Universal Robots URScript: test_first_drawing_!.script

def Machining1():
  # Default parameters:
  global speed_ms = 0.3
  global speed_rads = 0.75
  global accel_mss = 3
  global accel_radss = 1.2
  global blend_radius_m = 0.001

  # Add subprograms here
  # Start of main program
  # Program generated by RoboDK v5.6.5 for UR10e on 02/02/2024 16:16:45
  # Using nominal kinematics.
  blend_radius_m = 0.001
  speed_ms = 1.000
  # set_reference(p[0.123734, -0.255000, -0.004586, 0.000000, 0.000000, 0.000000])
  set_tcp(p[0.000000, 0.000000, 0.252000, 0.000000, 0.000000, 0.000000])
  # Show Tool
  movej([-0.457372, -0.718365, -2.572418, -1.421607, 1.570796, 1.113424],accel_radss,speed_rads,0,blend_radius_m)
  movel([-0.457372, -0.718365, -2.572418, -1.421607, 1.570796, 1.113424],accel_mss,speed_ms,0,blend_radius_m)
  # Splitting Linear movement in 6 (instruction 7: MoveL 3)
  movel([-0.457372, -0.726970, -2.600418, -1.385001, 1.570796, 1.113424],accel_mss,speed_ms,0,blend_radius_m)
  movel([-0.457372, -0.737986, -2.628172, -1.346232, 1.570796, 1.113424],accel_mss,speed_ms,0,blend_radius_m)
  movel([-0.457372, -0.751770, -2.655662, -1.304957, 1.570796, 1.113424],accel_mss,speed_ms,0,blend_radius_m)
  movel([-0.457372, -0.768751, -2.682869, -1.260769, 1.570796, 1.113424],accel_mss,speed_ms,0,blend_radius_m)
  movel([-0.457372, -0.789449, -2.709765, -1.213175, 1.570796, 1.113424],accel_mss,speed_ms,0,blend_radius_m)
  movel([-0.457372, -0.814491, -2.736314, -1.161584, 1.570796, 1.113424],accel_mss,speed_ms,0,blend_radius_m)
  movel([-0.457372, -0.814491, -2.736314, -1.161584, 1.570796, 1.113424],accel_mss,speed_ms,0,blend_radius_m)
  speed_ms = 1.000
  movel([-0.457372, -0.814491, -2.736314, -1.161584, 1.570796, 1.113424],accel_mss,speed_ms,0,blend_radius_m)
  movel([-0.457372, -0.814491, -2.736314, -1.161584, 1.570796, 1.113424],accel_mss,speed_ms,0,blend_radius_m)
  movel([-0.457372, -0.814491, -2.736314, -1.161584, 1.570796, 1.113424],accel_mss,speed_ms,0,blend_radius_m)
  speed_ms = 0.005
  movel([-0.457372, -0.784984, -2.704412, -1.222993, 1.570796, 1.113424],accel_mss,speed_ms,0,blend_radius_m)
  speed_ms = 1.000
  movel([-0.457372, -0.814491, -2.736314, -1.161584, 1.570796, 1.113424],accel_mss,speed_ms,0,blend_radius_m)
  speed_ms = 0.040
  movel([-0.457372, -0.814491, -2.736314, -1.161584, 1.570796, 1.113424],accel_mss,speed_ms,0,blend_radius_m)
  speed_ms = 1.000
  movel([-0.457372, -0.814491, -2.736314, -1.161584, 1.570796, 1.113424],accel_mss,speed_ms,0,blend_radius_m)
  # Splitting Linear movement in 8 (instruction 21: MoveL 12)
  movel([-0.394298, -0.800154, -2.739094, -1.173141, 1.570796, 1.176498],accel_mss,speed_ms,0,blend_radius_m)
  movel([-0.332487, -0.789840, -2.741023, -1.181526, 1.570796, 1.238309],accel_mss,speed_ms,0,blend_radius_m)
  movel([-0.272464, -0.783804, -2.742125, -1.186460, 1.570796, 1.298332],accel_mss,speed_ms,0,blend_radius_m)
  movel([-0.214704, -0.782203, -2.742414, -1.187772, 1.570796, 1.356092],accel_mss,speed_ms,0,blend_radius_m)
  movel([-0.159605, -0.785077, -2.741894, -1.185418, 1.570796, 1.411192],accel_mss,speed_ms,0,blend_radius_m)
  movel([-0.107470, -0.792353, -2.740559, -1.179478, 1.570796, 1.463327],accel_mss,speed_ms,0,blend_radius_m)
  movel([-0.058503, -0.803844, -2.738390, -1.170155, 1.570796, 1.512293],accel_mss,speed_ms,0,blend_radius_m)
  movel([-0.012808, -0.819267, -2.735362, -1.157760, 1.570796, 1.557988],accel_mss,speed_ms,0,blend_radius_m)
  speed_ms = 0.005
  movel([-0.012808, -0.856350, -2.766620, -1.089418, 1.570796, 1.557988],accel_mss,speed_ms,0,blend_radius_m)
  speed_ms = 0.025
  movel([-0.015705, -0.866064, -2.764578, -1.081748, 1.570796, 1.555091],accel_mss,speed_ms,0,blend_radius_m)
  movel([-0.017368, -0.870976, -2.763523, -1.077890, 1.570796, 1.553429],accel_mss,speed_ms,0,blend_radius_m)
  movel([-0.019216, -0.875915, -2.762449, -1.074025, 1.570796, 1.551580],accel_mss,speed_ms,0,blend_radius_m)
  movel([-0.021279, -0.880866, -2.761357, -1.070166, 1.570796, 1.549518],accel_mss,speed_ms,0,blend_radius_m)
  movel([-0.023584, -0.885818, -2.760249, -1.066321, 1.570796, 1.547213],accel_mss,speed_ms,0,blend_radius_m)
  movel([-0.026163, -0.890765, -2.759128, -1.062496, 1.570796, 1.544633],accel_mss,speed_ms,0,blend_radius_m)
  movel([-0.029049, -0.895692, -2.757997, -1.058701, 1.570796, 1.541747],accel_mss,speed_ms,0,blend_radius_m)
  movel([-0.028017, -0.893565, -2.758487, -1.060337, 1.570796, 1.542779],accel_mss,speed_ms,0,blend_radius_m)
  movel([-0.027153, -0.890950, -2.759086, -1.062353, 1.570796, 1.543644],accel_mss,speed_ms,0,blend_radius_m)
  movel([-0.026737, -0.888547, -2.759633, -1.064209, 1.570796, 1.544059],accel_mss,speed_ms,0,blend_radius_m)
  movel([-0.026791, -0.887653, -2.759835, -1.064900, 1.570796, 1.544006],accel_mss,speed_ms,0,blend_radius_m)
  movel([-0.027063, -0.887078, -2.759965, -1.065346, 1.570796, 1.543734],accel_mss,speed_ms,0,blend_radius_m)
  movel([-0.027595, -0.886898, -2.760006, -1.065485, 1.570796, 1.543202],accel_mss,speed_ms,0,blend_radius_m)
  movel([-0.028284, -0.887183, -2.759942, -1.065264, 1.570796, 1.542513],accel_mss,speed_ms,0,blend_radius_m)
  movel([-0.029095, -0.887869, -2.759787, -1.064734, 1.570796, 1.541701],accel_mss,speed_ms,0,blend_radius_m)
  movel([-0.030017, -0.888906, -2.759551, -1.063932, 1.570796, 1.540780],accel_mss,speed_ms,0,blend_radius_m)
  movel([-0.032071, -0.891780, -2.758896, -1.061712, 1.570796, 1.538725],accel_mss,speed_ms,0,blend_radius_m)
  movel([-0.034255, -0.895333, -2.758079, -1.058976, 1.570796, 1.536542],accel_mss,speed_ms,0,blend_radius_m)
  movel([-0.038281, -0.902664, -2.756369, -1.053356, 1.570796, 1.532515],accel_mss,speed_ms,0,blend_radius_m)
  movel([-0.040683, -0.907306, -2.755268, -1.049815, 1.570796, 1.530113],accel_mss,speed_ms,0,blend_radius_m)
  movel([-0.044313, -0.913830, -2.753697, -1.044862, 1.570796, 1.526483],accel_mss,speed_ms,0,blend_radius_m)
  movel([-0.046379, -0.916993, -2.752926, -1.042470, 1.570796, 1.524417],accel_mss,speed_ms,0,blend_radius_m)
  movel([-0.048725, -0.920005, -2.752185, -1.040199, 1.570796, 1.522072],accel_mss,speed_ms,0,blend_radius_m)
  movel([-0.048271, -0.919131, -2.752401, -1.040857, 1.570796, 1.522525],accel_mss,speed_ms,0,blend_radius_m)
  movel([-0.048029, -0.917919, -2.752699, -1.041771, 1.570796, 1.522767],accel_mss,speed_ms,0,blend_radius_m)
  movel([-0.048062, -0.915005, -2.753411, -1.043973, 1.570796, 1.522735],accel_mss,speed_ms,0,blend_radius_m)
  movel([-0.048591, -0.912345, -2.754057, -1.045987, 1.570796, 1.522205],accel_mss,speed_ms,0,blend_radius_m)
  movel([-0.048976, -0.911448, -2.754274, -1.046667, 1.570796, 1.521820],accel_mss,speed_ms,0,blend_radius_m)
  movel([-0.049395, -0.911024, -2.754376, -1.046989, 1.570796, 1.521401],accel_mss,speed_ms,0,blend_radius_m)
  movel([-0.050483, -0.910927, -2.754399, -1.047062, 1.570796, 1.520313],accel_mss,speed_ms,0,blend_radius_m)
  movel([-0.051522, -0.911310, -2.754307, -1.046772, 1.570796, 1.519275],accel_mss,speed_ms,0,blend_radius_m)
  movel([-0.052515, -0.912075, -2.754122, -1.046192, 1.570796, 1.518281],accel_mss,speed_ms,0,blend_radius_m)
  movel([-0.053463, -0.913130, -2.753867, -1.045392, 1.570796, 1.517333],accel_mss,speed_ms,0,blend_radius_m)
  movel([-0.055213, -0.915686, -2.753245, -1.043458, 1.570796, 1.515583],accel_mss,speed_ms,0,blend_radius_m)
  movel([-0.056771, -0.918197, -2.752631, -1.041562, 1.570796, 1.514025],accel_mss,speed_ms,0,blend_radius_m)
  movel([-0.059370, -0.922009, -2.751689, -1.038691, 1.570796, 1.511427],accel_mss,speed_ms,0,blend_radius_m)
  movel([-0.062062, -0.925527, -2.750812, -1.036050, 1.570796, 1.508735],accel_mss,speed_ms,0,blend_radius_m)
  movel([-0.065029, -0.928771, -2.749996, -1.033622, 1.570796, 1.505768],accel_mss,speed_ms,0,blend_radius_m)
  movel([-0.068441, -0.931736, -2.749244, -1.031409, 1.570796, 1.502355],accel_mss,speed_ms,0,blend_radius_m)
  movel([-0.066682, -0.928859, -2.749974, -1.033557, 1.570796, 1.504114],accel_mss,speed_ms,0,blend_radius_m)
  movel([-0.065327, -0.925996, -2.750694, -1.035699, 1.570796, 1.505469],accel_mss,speed_ms,0,blend_radius_m)
  movel([-0.064965, -0.924615, -2.751040, -1.036734, 1.570796, 1.505831],accel_mss,speed_ms,0,blend_radius_m)
  movel([-0.064915, -0.923396, -2.751344, -1.037649, 1.570796, 1.505881],accel_mss,speed_ms,0,blend_radius_m)
  movel([-0.065209, -0.922449, -2.751580, -1.038360, 1.570796, 1.505588],accel_mss,speed_ms,0,blend_radius_m)
  movel([-0.065897, -0.921914, -2.751713, -1.038762, 1.570796, 1.504899],accel_mss,speed_ms,0,blend_radius_m)
  movel([-0.067234, -0.921954, -2.751703, -1.038732, 1.570796, 1.503563],accel_mss,speed_ms,0,blend_radius_m)
  movel([-0.068837, -0.922643, -2.751532, -1.038214, 1.570796, 1.501959],accel_mss,speed_ms,0,blend_radius_m)
  movel([-0.070570, -0.923760, -2.751254, -1.037376, 1.570796, 1.500226],accel_mss,speed_ms,0,blend_radius_m)
  movel([-0.072285, -0.925061, -2.750929, -1.036399, 1.570796, 1.498511],accel_mss,speed_ms,0,blend_radius_m)
  speed_ms = 0.005
  movel([-0.072285, -0.916497, -2.744962, -1.050930, 1.570796, 1.498511],accel_mss,speed_ms,0,blend_radius_m)
  speed_ms = 0.040
  movel([-0.064341, -0.944955, -2.737631, -1.029804, 1.570796, 1.506455],accel_mss,speed_ms,0,blend_radius_m)
  speed_ms = 0.005
  movel([-0.064341, -0.953673, -2.743494, -1.015222, 1.570796, 1.506455],accel_mss,speed_ms,0,blend_radius_m)
  speed_ms = 0.025
  movel([-0.063744, -0.951411, -2.744102, -1.016876, 1.570796, 1.507052],accel_mss,speed_ms,0,blend_radius_m)
  movel([-0.062886, -0.949058, -2.744731, -1.018600, 1.570796, 1.507911],accel_mss,speed_ms,0,blend_radius_m)
  movel([-0.061790, -0.946658, -2.745368, -1.020363, 1.570796, 1.509006],accel_mss,speed_ms,0,blend_radius_m)
  movel([-0.060471, -0.944238, -2.746007, -1.022144, 1.570796, 1.510325],accel_mss,speed_ms,0,blend_radius_m)
  movel([-0.058951, -0.941831, -2.746638, -1.023920, 1.570796, 1.511845],accel_mss,speed_ms,0,blend_radius_m)
  movel([-0.057246, -0.939476, -2.747252, -1.025660, 1.570796, 1.513550],accel_mss,speed_ms,0,blend_radius_m)
  movel([-0.055380, -0.937209, -2.747840, -1.027340, 1.570796, 1.515416],accel_mss,speed_ms,0,blend_radius_m)
  movel([-0.053368, -0.935059, -2.748394, -1.028936, 1.570796, 1.517428],accel_mss,speed_ms,0,blend_radius_m)
  movel([-0.050202, -0.932150, -2.749138, -1.031101, 1.570796, 1.520594],accel_mss,speed_ms,0,blend_radius_m)
  movel([-0.047049, -0.929750, -2.749748, -1.032891, 1.570796, 1.523747],accel_mss,speed_ms,0,blend_radius_m)
  movel([-0.043926, -0.927829, -2.750233, -1.034326, 1.570796, 1.526870],accel_mss,speed_ms,0,blend_radius_m)
  movel([-0.040855, -0.926363, -2.750602, -1.035424, 1.570796, 1.529941],accel_mss,speed_ms,0,blend_radius_m)
  movel([-0.037852, -0.925322, -2.750863, -1.036204, 1.570796, 1.532944],accel_mss,speed_ms,0,blend_radius_m)
  movel([-0.034930, -0.924675, -2.751025, -1.036689, 1.570796, 1.535866],accel_mss,speed_ms,0,blend_radius_m)
  movel([-0.032111, -0.924395, -2.751095, -1.036899, 1.570796, 1.538685],accel_mss,speed_ms,0,blend_radius_m)
  movel([-0.029407, -0.924448, -2.751082, -1.036859, 1.570796, 1.541389],accel_mss,speed_ms,0,blend_radius_m)
  movel([-0.026834, -0.924800, -2.750994, -1.036595, 1.570796, 1.543962],accel_mss,speed_ms,0,blend_radius_m)
  movel([-0.024404, -0.925419, -2.750839, -1.036131, 1.570796, 1.546392],accel_mss,speed_ms,0,blend_radius_m)
  movel([-0.020023, -0.927315, -2.750363, -1.034711, 1.570796, 1.550774],accel_mss,speed_ms,0,blend_radius_m)
  movel([-0.016359, -0.929848, -2.749723, -1.032818, 1.570796, 1.554437],accel_mss,speed_ms,0,blend_radius_m)
  movel([-0.013508, -0.932744, -2.748987, -1.030659, 1.570796, 1.557288],accel_mss,speed_ms,0,blend_radius_m)
  movel([-0.011055, -0.936237, -2.748091, -1.028061, 1.570796, 1.559741],accel_mss,speed_ms,0,blend_radius_m)
  movel([-0.009001, -0.940105, -2.747089, -1.025195, 1.570796, 1.561795],accel_mss,speed_ms,0,blend_radius_m)
  movel([-0.007301, -0.944288, -2.745994, -1.022107, 1.570796, 1.563495],accel_mss,speed_ms,0,blend_radius_m)
  movel([-0.005915, -0.948731, -2.744818, -1.018840, 1.570796, 1.564881],accel_mss,speed_ms,0,blend_radius_m)
  movel([-0.004799, -0.953378, -2.743573, -1.015438, 1.570796, 1.565997],accel_mss,speed_ms,0,blend_radius_m)
  movel([-0.003906, -0.958173, -2.742273, -1.011943, 1.570796, 1.566890],accel_mss,speed_ms,0,blend_radius_m)
  movel([-0.002624, -0.967997, -2.739559, -1.004833, 1.570796, 1.568172],accel_mss,speed_ms,0,blend_radius_m)
  movel([-0.001812, -0.974866, -2.737620, -0.999903, 1.570796, 1.568984],accel_mss,speed_ms,0,blend_radius_m)
  movel([-0.001114, -0.978051, -2.736709, -0.997629, 1.570796, 1.569682],accel_mss,speed_ms,0,blend_radius_m)
  movel([-0.000027, -0.980907, -2.735886, -0.995596, 1.570796, 1.570769],accel_mss,speed_ms,0,blend_radius_m)
  movel([0.001984, -0.984157, -2.734942, -0.993289, 1.570796, 1.572780],accel_mss,speed_ms,0,blend_radius_m)
  movel([0.003993, -0.987421, -2.733987, -0.990981, 1.570796, 1.574789],accel_mss,speed_ms,0,blend_radius_m)
  movel([0.004723, -0.989213, -2.733459, -0.989717, 1.570796, 1.575519],accel_mss,speed_ms,0,blend_radius_m)
  movel([0.005120, -0.991196, -2.732872, -0.988321, 1.570796, 1.575917],accel_mss,speed_ms,0,blend_radius_m)
  movel([0.005081, -0.993422, -2.732209, -0.986758, 1.570796, 1.575877],accel_mss,speed_ms,0,blend_radius_m)
  movel([0.004502, -0.995954, -2.731451, -0.984984, 1.570796, 1.575298],accel_mss,speed_ms,0,blend_radius_m)
  movel([0.006531, -0.989512, -2.733371, -0.989507, 1.570796, 1.577327],accel_mss,speed_ms,0,blend_radius_m)
  movel([0.008255, -0.983151, -2.735235, -0.994002, 1.570796, 1.579051],accel_mss,speed_ms,0,blend_radius_m)
  movel([0.011148, -0.970478, -2.738862, -1.003048, 1.570796, 1.581944],accel_mss,speed_ms,0,blend_radius_m)
  movel([0.012546, -0.963426, -2.740830, -1.008133, 1.570796, 1.583343],accel_mss,speed_ms,0,blend_radius_m)
  movel([0.013759, -0.956404, -2.742755, -1.013230, 1.570796, 1.584556],accel_mss,speed_ms,0,blend_radius_m)
  movel([0.015756, -0.942395, -2.746491, -1.023503, 1.570796, 1.586553],accel_mss,speed_ms,0,blend_radius_m)
  movel([0.017248, -0.928713, -2.750010, -1.033665, 1.570796, 1.588045],accel_mss,speed_ms,0,blend_radius_m)
  movel([0.017651, -0.921969, -2.751699, -1.038721, 1.570796, 1.588447],accel_mss,speed_ms,0,blend_radius_m)
  movel([0.017671, -0.915464, -2.753299, -1.043625, 1.570796, 1.588467],accel_mss,speed_ms,0,blend_radius_m)
  movel([0.017291, -0.910583, -2.754482, -1.047323, 1.570796, 1.588087],accel_mss,speed_ms,0,blend_radius_m)
  movel([0.016655, -0.905838, -2.755617, -1.050933, 1.570796, 1.587451],accel_mss,speed_ms,0,blend_radius_m)
  movel([0.016029, -0.901034, -2.756752, -1.054603, 1.570796, 1.586825],accel_mss,speed_ms,0,blend_radius_m)
  movel([0.015681, -0.895972, -2.757932, -1.058485, 1.570796, 1.586478],accel_mss,speed_ms,0,blend_radius_m)
  movel([0.015770, -0.894507, -2.758270, -1.059612, 1.570796, 1.586566],accel_mss,speed_ms,0,blend_radius_m)
  movel([0.016153, -0.892883, -2.758644, -1.060862, 1.570796, 1.586949],accel_mss,speed_ms,0,blend_radius_m)
  movel([0.016912, -0.891306, -2.759005, -1.062078, 1.570796, 1.587708],accel_mss,speed_ms,0,blend_radius_m)
  movel([0.017466, -0.890591, -2.759168, -1.062630, 1.570796, 1.588262],accel_mss,speed_ms,0,blend_radius_m)
  movel([0.018150, -0.889955, -2.759313, -1.063121, 1.570796, 1.588946],accel_mss,speed_ms,0,blend_radius_m)
  movel([0.019160, -0.889356, -2.759449, -1.063583, 1.570796, 1.589956],accel_mss,speed_ms,0,blend_radius_m)
  movel([0.020130, -0.889010, -2.759528, -1.063851, 1.570796, 1.590927],accel_mss,speed_ms,0,blend_radius_m)
  movel([0.025280, -0.887760, -2.759811, -1.064818, 1.570796, 1.596076],accel_mss,speed_ms,0,blend_radius_m)
  movel([0.029950, -0.887246, -2.759927, -1.065216, 1.570796, 1.600746],accel_mss,speed_ms,0,blend_radius_m)
  movel([0.034170, -0.887403, -2.759892, -1.065094, 1.570796, 1.604966],accel_mss,speed_ms,0,blend_radius_m)
  movel([0.037971, -0.888183, -2.759715, -1.064490, 1.570796, 1.608767],accel_mss,speed_ms,0,blend_radius_m)
  movel([0.041380, -0.889522, -2.759412, -1.063456, 1.570796, 1.612176],accel_mss,speed_ms,0,blend_radius_m)
  movel([0.044433, -0.891356, -2.758993, -1.062040, 1.570796, 1.615229],accel_mss,speed_ms,0,blend_radius_m)
  movel([0.047160, -0.893627, -2.758473, -1.060289, 1.570796, 1.617956],accel_mss,speed_ms,0,blend_radius_m)
  movel([0.049593, -0.896280, -2.757860, -1.058249, 1.570796, 1.620390],accel_mss,speed_ms,0,blend_radius_m)
  movel([0.051770, -0.899248, -2.757170, -1.055971, 1.570796, 1.622566],accel_mss,speed_ms,0,blend_radius_m)
  movel([0.053728, -0.902471, -2.756414, -1.053504, 1.570796, 1.624524],accel_mss,speed_ms,0,blend_radius_m)
  movel([0.057117, -0.909448, -2.754755, -1.048186, 1.570796, 1.627913],accel_mss,speed_ms,0,blend_radius_m)
  movel([0.062777, -0.923949, -2.751206, -1.037234, 1.570796, 1.633573],accel_mss,speed_ms,0,blend_radius_m)
  movel([0.063800, -0.926089, -2.750671, -1.035629, 1.570796, 1.634597],accel_mss,speed_ms,0,blend_radius_m)
  movel([0.064540, -0.926900, -2.750467, -1.035021, 1.570796, 1.635337],accel_mss,speed_ms,0,blend_radius_m)
  movel([0.065528, -0.927402, -2.750341, -1.034646, 1.570796, 1.636324],accel_mss,speed_ms,0,blend_radius_m)
  movel([0.067440, -0.927423, -2.750336, -1.034630, 1.570796, 1.638236],accel_mss,speed_ms,0,blend_radius_m)
  movel([0.068455, -0.927126, -2.750410, -1.034852, 1.570796, 1.639251],accel_mss,speed_ms,0,blend_radius_m)
  movel([0.069499, -0.926643, -2.750532, -1.035214, 1.570796, 1.640295],accel_mss,speed_ms,0,blend_radius_m)
  movel([0.071627, -0.925216, -2.750890, -1.036283, 1.570796, 1.642424],accel_mss,speed_ms,0,blend_radius_m)
  movel([0.073755, -0.923294, -2.751370, -1.037725, 1.570796, 1.644551],accel_mss,speed_ms,0,blend_radius_m)
  movel([0.075801, -0.921041, -2.751929, -1.039419, 1.570796, 1.646597],accel_mss,speed_ms,0,blend_radius_m)
  movel([0.077686, -0.918613, -2.752528, -1.041247, 1.570796, 1.648483],accel_mss,speed_ms,0,blend_radius_m)
  movel([0.079336, -0.916165, -2.753128, -1.043095, 1.570796, 1.650133],accel_mss,speed_ms,0,blend_radius_m)
  movel([0.080656, -0.913866, -2.753688, -1.044834, 1.570796, 1.651452],accel_mss,speed_ms,0,blend_radius_m)
  movel([0.082630, -0.909930, -2.754640, -1.047820, 1.570796, 1.653426],accel_mss,speed_ms,0,blend_radius_m)
  movel([0.084460, -0.905965, -2.755587, -1.050837, 1.570796, 1.655256],accel_mss,speed_ms,0,blend_radius_m)
  movel([0.087673, -0.898016, -2.757457, -1.056916, 1.570796, 1.658469],accel_mss,speed_ms,0,blend_radius_m)
  movel([0.090296, -0.890146, -2.759269, -1.062974, 1.570796, 1.661093],accel_mss,speed_ms,0,blend_radius_m)
  movel([0.092317, -0.882486, -2.760996, -1.068906, 1.570796, 1.663113],accel_mss,speed_ms,0,blend_radius_m)
  movel([0.092972, -0.879636, -2.761629, -1.071123, 1.570796, 1.663768],accel_mss,speed_ms,0,blend_radius_m)
  movel([0.093861, -0.876714, -2.762274, -1.073401, 1.570796, 1.664657],accel_mss,speed_ms,0,blend_radius_m)
  movel([0.094496, -0.875233, -2.762598, -1.074558, 1.570796, 1.665293],accel_mss,speed_ms,0,blend_radius_m)
  movel([0.095316, -0.873730, -2.762926, -1.075733, 1.570796, 1.666112],accel_mss,speed_ms,0,blend_radius_m)
  movel([0.096359, -0.872215, -2.763255, -1.076919, 1.570796, 1.667155],accel_mss,speed_ms,0,blend_radius_m)
  movel([0.097667, -0.870690, -2.763585, -1.078114, 1.570796, 1.668463],accel_mss,speed_ms,0,blend_radius_m)
  movel([0.099645, -0.869011, -2.763947, -1.079431, 1.570796, 1.670442],accel_mss,speed_ms,0,blend_radius_m)
  movel([0.101657, -0.867976, -2.764169, -1.080244, 1.570796, 1.672454],accel_mss,speed_ms,0,blend_radius_m)
  movel([0.103554, -0.867531, -2.764264, -1.080594, 1.570796, 1.674351],accel_mss,speed_ms,0,blend_radius_m)
  movel([0.105201, -0.867609, -2.764248, -1.080532, 1.570796, 1.675998],accel_mss,speed_ms,0,blend_radius_m)
  movel([0.107545, -0.868375, -2.764083, -1.079931, 1.570796, 1.678341],accel_mss,speed_ms,0,blend_radius_m)
  movel([0.109640, -0.869541, -2.763833, -1.079015, 1.570796, 1.680436],accel_mss,speed_ms,0,blend_radius_m)
  movel([0.113241, -0.872557, -2.763181, -1.076651, 1.570796, 1.684037],accel_mss,speed_ms,0,blend_radius_m)
  movel([0.114694, -0.874237, -2.762816, -1.075336, 1.570796, 1.685491],accel_mss,speed_ms,0,blend_radius_m)
  movel([0.115871, -0.876122, -2.762404, -1.073864, 1.570796, 1.686668],accel_mss,speed_ms,0,blend_radius_m)
  movel([0.116792, -0.878190, -2.761949, -1.072250, 1.570796, 1.687588],accel_mss,speed_ms,0,blend_radius_m)
  movel([0.117465, -0.880433, -2.761453, -1.070503, 1.570796, 1.688262],accel_mss,speed_ms,0,blend_radius_m)
  movel([0.117909, -0.882834, -2.760919, -1.068636, 1.570796, 1.688705],accel_mss,speed_ms,0,blend_radius_m)
  movel([0.118158, -0.888067, -2.759742, -1.064581, 1.570796, 1.688954],accel_mss,speed_ms,0,blend_radius_m)
  movel([0.117990, -0.890869, -2.759105, -1.062415, 1.570796, 1.688786],accel_mss,speed_ms,0,blend_radius_m)
  movel([0.117154, -0.896775, -2.757746, -1.057869, 1.570796, 1.687950],accel_mss,speed_ms,0,blend_radius_m)
  movel([0.115733, -0.903003, -2.756289, -1.053097, 1.570796, 1.686529],accel_mss,speed_ms,0,blend_radius_m)
  movel([0.113833, -0.909462, -2.754752, -1.048175, 1.570796, 1.684629],accel_mss,speed_ms,0,blend_radius_m)
  movel([0.111569, -0.916046, -2.753158, -1.043186, 1.570796, 1.682366],accel_mss,speed_ms,0,blend_radius_m)
  movel([0.107783, -0.925727, -2.750762, -1.035900, 1.570796, 1.678579],accel_mss,speed_ms,0,blend_radius_m)
  movel([0.105653, -0.930585, -2.749536, -1.032268, 1.570796, 1.676449],accel_mss,speed_ms,0,blend_radius_m)
  movel([0.103334, -0.935430, -2.748298, -1.028661, 1.570796, 1.674131],accel_mss,speed_ms,0,blend_radius_m)
  movel([0.100810, -0.940237, -2.747054, -1.025097, 1.570796, 1.671606],accel_mss,speed_ms,0,blend_radius_m)
  movel([0.098064, -0.944987, -2.745810, -1.021592, 1.570796, 1.668860],accel_mss,speed_ms,0,blend_radius_m)
  movel([0.095066, -0.949669, -2.744568, -1.018152, 1.570796, 1.665862],accel_mss,speed_ms,0,blend_radius_m)
  movel([0.091805, -0.954256, -2.743336, -1.014797, 1.570796, 1.662601],accel_mss,speed_ms,0,blend_radius_m)
  movel([0.086890, -0.960481, -2.741642, -1.010267, 1.570796, 1.657687],accel_mss,speed_ms,0,blend_radius_m)
  movel([0.084158, -0.963622, -2.740776, -1.007991, 1.570796, 1.654954],accel_mss,speed_ms,0,blend_radius_m)
  movel([0.081297, -0.966623, -2.739942, -1.005824, 1.570796, 1.652094],accel_mss,speed_ms,0,blend_radius_m)
  movel([0.078356, -0.969360, -2.739177, -1.003852, 1.570796, 1.649152],accel_mss,speed_ms,0,blend_radius_m)
  movel([0.075374, -0.971717, -2.738513, -1.002159, 1.570796, 1.646170],accel_mss,speed_ms,0,blend_radius_m)
  movel([0.072391, -0.973574, -2.737987, -1.000828, 1.570796, 1.643187],accel_mss,speed_ms,0,blend_radius_m)
  movel([0.070913, -0.974281, -2.737786, -1.000322, 1.570796, 1.641710],accel_mss,speed_ms,0,blend_radius_m)
  movel([0.069453, -0.974815, -2.737634, -0.999940, 1.570796, 1.640249],accel_mss,speed_ms,0,blend_radius_m)
  movel([0.067859, -0.975193, -2.737527, -0.999670, 1.570796, 1.638655],accel_mss,speed_ms,0,blend_radius_m)
  movel([0.066391, -0.975318, -2.737491, -0.999580, 1.570796, 1.637187],accel_mss,speed_ms,0,blend_radius_m)
  movel([0.065038, -0.975217, -2.737520, -0.999652, 1.570796, 1.635834],accel_mss,speed_ms,0,blend_radius_m)
  movel([0.063796, -0.974907, -2.737608, -0.999874, 1.570796, 1.634592],accel_mss,speed_ms,0,blend_radius_m)
  movel([0.061607, -0.973759, -2.737935, -1.000696, 1.570796, 1.632403],accel_mss,speed_ms,0,blend_radius_m)
  movel([0.059773, -0.972041, -2.738421, -1.001927, 1.570796, 1.630570],accel_mss,speed_ms,0,blend_radius_m)
  movel([0.058238, -0.969934, -2.739015, -1.003440, 1.570796, 1.629034],accel_mss,speed_ms,0,blend_radius_m)
  movel([0.056949, -0.967612, -2.739666, -1.005111, 1.570796, 1.627745],accel_mss,speed_ms,0,blend_radius_m)
  movel([0.054905, -0.963026, -2.740941, -1.008422, 1.570796, 1.625701],accel_mss,speed_ms,0,blend_radius_m)
  movel([0.053979, -0.960865, -2.741536, -1.009988, 1.570796, 1.624775],accel_mss,speed_ms,0,blend_radius_m)
  movel([0.052794, -0.958972, -2.742055, -1.011362, 1.570796, 1.623591],accel_mss,speed_ms,0,blend_radius_m)
  movel([0.051998, -0.958284, -2.742243, -1.011862, 1.570796, 1.622794],accel_mss,speed_ms,0,blend_radius_m)
  movel([0.051005, -0.957852, -2.742361, -1.012176, 1.570796, 1.621801],accel_mss,speed_ms,0,blend_radius_m)
  movel([0.049778, -0.957741, -2.742391, -1.012257, 1.570796, 1.620574],accel_mss,speed_ms,0,blend_radius_m)
  movel([0.048272, -0.958009, -2.742318, -1.012062, 1.570796, 1.619069],accel_mss,speed_ms,0,blend_radius_m)
  movel([0.048603, -0.958015, -2.742316, -1.012058, 1.570796, 1.619399],accel_mss,speed_ms,0,blend_radius_m)
  movel([0.048805, -0.958251, -2.742252, -1.011886, 1.570796, 1.619602],accel_mss,speed_ms,0,blend_radius_m)
  movel([0.048847, -0.959360, -2.741949, -1.011080, 1.570796, 1.619643],accel_mss,speed_ms,0,blend_radius_m)
  movel([0.048450, -0.961220, -2.741439, -1.009731, 1.570796, 1.619246],accel_mss,speed_ms,0,blend_radius_m)
  movel([0.047686, -0.963709, -2.740752, -1.007928, 1.570796, 1.618482],accel_mss,speed_ms,0,blend_radius_m)
  movel([0.045299, -0.970090, -2.738971, -1.003327, 1.570796, 1.616095],accel_mss,speed_ms,0,blend_radius_m)
  movel([0.042178, -0.977549, -2.736853, -0.997987, 1.570796, 1.612974],accel_mss,speed_ms,0,blend_radius_m)
  movel([0.035644, -0.992051, -2.732618, -0.987721, 1.570796, 1.606440],accel_mss,speed_ms,0,blend_radius_m)
  movel([0.031683, -1.000255, -2.730152, -0.981982, 1.570796, 1.602480],accel_mss,speed_ms,0,blend_radius_m)
  movel([0.026965, -1.008739, -2.727549, -0.976102, 1.570796, 1.597761],accel_mss,speed_ms,0,blend_radius_m)
  movel([0.022176, -1.017023, -2.724953, -0.970413, 1.570796, 1.592972],accel_mss,speed_ms,0,blend_radius_m)
  movel([0.017300, -1.025189, -2.722341, -0.964859, 1.570796, 1.588096],accel_mss,speed_ms,0,blend_radius_m)
  movel([0.007614, -1.040765, -2.717211, -0.954413, 1.570796, 1.578410],accel_mss,speed_ms,0,blend_radius_m)
  movel([0.002683, -1.048049, -2.714744, -0.949595, 1.570796, 1.573479],accel_mss,speed_ms,0,blend_radius_m)
  movel([0.000072, -1.051561, -2.713539, -0.947289, 1.570796, 1.570868],accel_mss,speed_ms,0,blend_radius_m)
  movel([-0.002659, -1.054953, -2.712365, -0.945071, 1.570796, 1.568137],accel_mss,speed_ms,0,blend_radius_m)
  movel([-0.005542, -1.058200, -2.711233, -0.942956, 1.570796, 1.565254],accel_mss,speed_ms,0,blend_radius_m)
  movel([-0.008588, -1.061277, -2.710151, -0.940961, 1.570796, 1.562208],accel_mss,speed_ms,0,blend_radius_m)
  movel([-0.008300, -1.055649, -2.712123, -0.944617, 1.570796, 1.562497],accel_mss,speed_ms,0,blend_radius_m)
  movel([-0.008450, -1.054105, -2.712660, -0.945624, 1.570796, 1.562346],accel_mss,speed_ms,0,blend_radius_m)
  movel([-0.008799, -1.053604, -2.712833, -0.945952, 1.570796, 1.561997],accel_mss,speed_ms,0,blend_radius_m)
  movel([-0.009432, -1.053476, -2.712878, -0.946035, 1.570796, 1.561364],accel_mss,speed_ms,0,blend_radius_m)
  movel([-0.010104, -1.053708, -2.712797, -0.945883, 1.570796, 1.560692],accel_mss,speed_ms,0,blend_radius_m)
  movel([-0.010802, -1.054169, -2.712638, -0.945583, 1.570796, 1.559994],accel_mss,speed_ms,0,blend_radius_m)
  movel([-0.014070, -1.056982, -2.711659, -0.943748, 1.570796, 1.556726],accel_mss,speed_ms,0,blend_radius_m)
  movel([-0.016026, -1.058338, -2.711184, -0.942867, 1.570796, 1.554770],accel_mss,speed_ms,0,blend_radius_m)
  movel([-0.018005, -1.059430, -2.710801, -0.942158, 1.570796, 1.552792],accel_mss,speed_ms,0,blend_radius_m)
  movel([-0.019956, -1.060230, -2.710520, -0.941639, 1.570796, 1.550841],accel_mss,speed_ms,0,blend_radius_m)
  movel([-0.020553, -1.060316, -2.710490, -0.941583, 1.570796, 1.550244],accel_mss,speed_ms,0,blend_radius_m)
  movel([-0.020750, -1.060021, -2.710594, -0.941775, 1.570796, 1.550047],accel_mss,speed_ms,0,blend_radius_m)
  movel([-0.020330, -1.058298, -2.711198, -0.942893, 1.570796, 1.550466],accel_mss,speed_ms,0,blend_radius_m)
  movel([-0.020427, -1.057821, -2.711365, -0.943202, 1.570796, 1.550369],accel_mss,speed_ms,0,blend_radius_m)
  movel([-0.020779, -1.057569, -2.711454, -0.943367, 1.570796, 1.550018],accel_mss,speed_ms,0,blend_radius_m)
  movel([-0.021298, -1.057529, -2.711467, -0.943393, 1.570796, 1.549498],accel_mss,speed_ms,0,blend_radius_m)
  movel([-0.021902, -1.057693, -2.711410, -0.943286, 1.570796, 1.548894],accel_mss,speed_ms,0,blend_radius_m)
  movel([-0.023143, -1.058460, -2.711142, -0.942788, 1.570796, 1.547654],accel_mss,speed_ms,0,blend_radius_m)
  movel([-0.031654, -1.066064, -2.708452, -0.937873, 1.570796, 1.539142],accel_mss,speed_ms,0,blend_radius_m)
  movel([-0.029187, -1.063378, -2.709408, -0.939603, 1.570796, 1.541609],accel_mss,speed_ms,0,blend_radius_m)
  movel([-0.026775, -1.060512, -2.710421, -0.941457, 1.570796, 1.544022],accel_mss,speed_ms,0,blend_radius_m)
  movel([-0.024437, -1.057512, -2.711473, -0.943404, 1.570796, 1.546359],accel_mss,speed_ms,0,blend_radius_m)
  movel([-0.022179, -1.054410, -2.712554, -0.945425, 1.570796, 1.548617],accel_mss,speed_ms,0,blend_radius_m)
  movel([-0.017959, -1.048048, -2.714745, -0.949597, 1.570796, 1.552837],accel_mss,speed_ms,0,blend_radius_m)
  movel([-0.014223, -1.041744, -2.716882, -0.953763, 1.570796, 1.556573],accel_mss,speed_ms,0,blend_radius_m)
  movel([-0.010453, -1.034858, -2.719180, -0.958352, 1.570796, 1.560343],accel_mss,speed_ms,0,blend_radius_m)
  movel([-0.006899, -1.027854, -2.721477, -0.963057, 1.570796, 1.563897],accel_mss,speed_ms,0,blend_radius_m)
  movel([-0.005272, -1.024335, -2.722617, -0.965438, 1.570796, 1.565524],accel_mss,speed_ms,0,blend_radius_m)
  movel([-0.003775, -1.020815, -2.723747, -0.967828, 1.570796, 1.567021],accel_mss,speed_ms,0,blend_radius_m)
  movel([-0.002443, -1.017311, -2.724861, -0.970216, 1.570796, 1.568354],accel_mss,speed_ms,0,blend_radius_m)
  movel([-0.001298, -1.013828, -2.725960, -0.972601, 1.570796, 1.569498],accel_mss,speed_ms,0,blend_radius_m)
  movel([-0.000737, -1.011694, -2.726629, -0.974066, 1.570796, 1.570060],accel_mss,speed_ms,0,blend_radius_m)
  movel([-0.000345, -1.009600, -2.727281, -0.975507, 1.570796, 1.570452],accel_mss,speed_ms,0,blend_radius_m)
  movel([-0.000026, -1.005553, -2.728533, -0.978303, 1.570796, 1.570770],accel_mss,speed_ms,0,blend_radius_m)
  movel([-0.000280, -1.001733, -2.729702, -0.980953, 1.570796, 1.570517],accel_mss,speed_ms,0,blend_radius_m)
  movel([-0.001044, -0.998182, -2.730780, -0.983427, 1.570796, 1.569752],accel_mss,speed_ms,0,blend_radius_m)
  movel([-0.002245, -0.994936, -2.731756, -0.985696, 1.570796, 1.568551],accel_mss,speed_ms,0,blend_radius_m)
  movel([-0.003811, -0.992035, -2.732623, -0.987732, 1.570796, 1.566986],accel_mss,speed_ms,0,blend_radius_m)
  movel([-0.005678, -0.989521, -2.733368, -0.989500, 1.570796, 1.565118],accel_mss,speed_ms,0,blend_radius_m)
  movel([-0.007767, -0.987427, -2.733985, -0.990977, 1.570796, 1.563029],accel_mss,speed_ms,0,blend_radius_m)
  movel([-0.009278, -0.986640, -2.734216, -0.991533, 1.570796, 1.561518],accel_mss,speed_ms,0,blend_radius_m)
  movel([-0.011068, -0.986527, -2.734249, -0.991612, 1.570796, 1.559729],accel_mss,speed_ms,0,blend_radius_m)
  movel([-0.013033, -0.987029, -2.734102, -0.991258, 1.570796, 1.557763],accel_mss,speed_ms,0,blend_radius_m)
  movel([-0.015068, -0.988082, -2.733793, -0.990515, 1.570796, 1.555729],accel_mss,speed_ms,0,blend_radius_m)
  movel([-0.017075, -0.989619, -2.733339, -0.989431, 1.570796, 1.553721],accel_mss,speed_ms,0,blend_radius_m)
  movel([-0.018953, -0.991579, -2.732758, -0.988052, 1.570796, 1.551843],accel_mss,speed_ms,0,blend_radius_m)
  movel([-0.020593, -0.993887, -2.732070, -0.986432, 1.570796, 1.550204],accel_mss,speed_ms,0,blend_radius_m)
  movel([-0.021902, -0.996480, -2.731293, -0.984616, 1.570796, 1.548895],accel_mss,speed_ms,0,blend_radius_m)
  movel([-0.023588, -1.000418, -2.730103, -0.981868, 1.570796, 1.547208],accel_mss,speed_ms,0,blend_radius_m)
  movel([-0.025438, -1.004334, -2.728907, -0.979148, 1.570796, 1.545359],accel_mss,speed_ms,0,blend_radius_m)
  movel([-0.027473, -1.008197, -2.727717, -0.976475, 1.570796, 1.543323],accel_mss,speed_ms,0,blend_radius_m)
  movel([-0.029724, -1.011987, -2.726537, -0.973865, 1.570796, 1.541072],accel_mss,speed_ms,0,blend_radius_m)
  movel([-0.032206, -1.015673, -2.725380, -0.971337, 1.570796, 1.538590],accel_mss,speed_ms,0,blend_radius_m)
  movel([-0.034949, -1.019235, -2.724251, -0.968904, 1.570796, 1.535847],accel_mss,speed_ms,0,blend_radius_m)
  movel([-0.037977, -1.022651, -2.723158, -0.966579, 1.570796, 1.532820],accel_mss,speed_ms,0,blend_radius_m)
  movel([-0.041308, -1.025896, -2.722112, -0.964381, 1.570796, 1.529489],accel_mss,speed_ms,0,blend_radius_m)
  movel([-0.043141, -1.027404, -2.721623, -0.963361, 1.570796, 1.527656],accel_mss,speed_ms,0,blend_radius_m)
  movel([-0.045025, -1.028711, -2.721198, -0.962480, 1.570796, 1.525771],accel_mss,speed_ms,0,blend_radius_m)
  movel([-0.048851, -1.030951, -2.720466, -0.960972, 1.570796, 1.521945],accel_mss,speed_ms,0,blend_radius_m)
  movel([-0.051855, -1.032427, -2.719982, -0.959980, 1.570796, 1.518942],accel_mss,speed_ms,0,blend_radius_m)
  movel([-0.054729, -1.033492, -2.719631, -0.959266, 1.570796, 1.516067],accel_mss,speed_ms,0,blend_radius_m)
  movel([-0.057472, -1.034176, -2.719405, -0.958808, 1.570796, 1.513324],accel_mss,speed_ms,0,blend_radius_m)
  movel([-0.060093, -1.034512, -2.719294, -0.958583, 1.570796, 1.510703],accel_mss,speed_ms,0,blend_radius_m)
  movel([-0.062595, -1.034534, -2.719287, -0.958568, 1.570796, 1.508201],accel_mss,speed_ms,0,blend_radius_m)
  movel([-0.064982, -1.034272, -2.719374, -0.958744, 1.570796, 1.505814],accel_mss,speed_ms,0,blend_radius_m)
  movel([-0.067250, -1.033750, -2.719546, -0.959093, 1.570796, 1.503546],accel_mss,speed_ms,0,blend_radius_m)
  movel([-0.069405, -1.033003, -2.719792, -0.959594, 1.570796, 1.501391],accel_mss,speed_ms,0,blend_radius_m)
  movel([-0.071449, -1.032061, -2.720102, -0.960226, 1.570796, 1.499347],accel_mss,speed_ms,0,blend_radius_m)
  movel([-0.073381, -1.030945, -2.720468, -0.960975, 1.570796, 1.497415],accel_mss,speed_ms,0,blend_radius_m)
  movel([-0.076913, -1.028330, -2.721322, -0.962736, 1.570796, 1.493884],accel_mss,speed_ms,0,blend_radius_m)
  movel([-0.080004, -1.025382, -2.722279, -0.964728, 1.570796, 1.490792],accel_mss,speed_ms,0,blend_radius_m)
  movel([-0.082651, -1.022337, -2.723259, -0.966793, 1.570796, 1.488146],accel_mss,speed_ms,0,blend_radius_m)
  movel([-0.084495, -1.019837, -2.724059, -0.968493, 1.570796, 1.486301],accel_mss,speed_ms,0,blend_radius_m)
  movel([-0.086208, -1.017088, -2.724932, -0.970369, 1.570796, 1.484589],accel_mss,speed_ms,0,blend_radius_m)
  movel([-0.087768, -1.014096, -2.725876, -0.972417, 1.570796, 1.483028],accel_mss,speed_ms,0,blend_radius_m)
  movel([-0.089137, -1.010871, -2.726886, -0.974632, 1.570796, 1.481659],accel_mss,speed_ms,0,blend_radius_m)
  movel([-0.090297, -1.007423, -2.727956, -0.977010, 1.570796, 1.480500],accel_mss,speed_ms,0,blend_radius_m)
  movel([-0.091211, -1.003760, -2.729083, -0.979546, 1.570796, 1.479586],accel_mss,speed_ms,0,blend_radius_m)
  movel([-0.091847, -0.999887, -2.730264, -0.982238, 1.570796, 1.478949],accel_mss,speed_ms,0,blend_radius_m)
  movel([-0.092176, -0.995812, -2.731494, -0.985083, 1.570796, 1.478621],accel_mss,speed_ms,0,blend_radius_m)
  movel([-0.092167, -0.991541, -2.732769, -0.988079, 1.570796, 1.478629],accel_mss,speed_ms,0,blend_radius_m)
  movel([-0.091786, -0.987087, -2.734085, -0.991217, 1.570796, 1.479010],accel_mss,speed_ms,0,blend_radius_m)
  movel([-0.091001, -0.982448, -2.735440, -0.994501, 1.570796, 1.479795],accel_mss,speed_ms,0,blend_radius_m)
  movel([-0.089771, -0.977635, -2.736828, -0.997926, 1.570796, 1.481025],accel_mss,speed_ms,0,blend_radius_m)
  movel([-0.088067, -0.972657, -2.738247, -1.001485, 1.570796, 1.482729],accel_mss,speed_ms,0,blend_radius_m)
  movel([-0.085849, -0.967515, -2.739693, -1.005180, 1.570796, 1.484947],accel_mss,speed_ms,0,blend_radius_m)
  movel([-0.083084, -0.962228, -2.741161, -1.009000, 1.570796, 1.487712],accel_mss,speed_ms,0,blend_radius_m)
  movel([-0.079736, -0.956800, -2.742647, -1.012942, 1.570796, 1.491060],accel_mss,speed_ms,0,blend_radius_m)
  movel([-0.078244, -0.954732, -2.743208, -1.014449, 1.570796, 1.492552],accel_mss,speed_ms,0,blend_radius_m)
  movel([-0.077402, -0.953783, -2.743464, -1.015142, 1.570796, 1.493394],accel_mss,speed_ms,0,blend_radius_m)
  movel([-0.076483, -0.952964, -2.743685, -1.015741, 1.570796, 1.494314],accel_mss,speed_ms,0,blend_radius_m)
  movel([-0.075051, -0.952139, -2.743907, -1.016344, 1.570796, 1.495745],accel_mss,speed_ms,0,blend_radius_m)
  movel([-0.073726, -0.951837, -2.743988, -1.016564, 1.570796, 1.497071],accel_mss,speed_ms,0,blend_radius_m)
  movel([-0.072569, -0.951977, -2.743950, -1.016462, 1.570796, 1.498227],accel_mss,speed_ms,0,blend_radius_m)
  movel([-0.071650, -0.952476, -2.743816, -1.016097, 1.570796, 1.499146],accel_mss,speed_ms,0,blend_radius_m)
  movel([-0.070227, -0.954257, -2.743336, -1.014796, 1.570796, 1.500570],accel_mss,speed_ms,0,blend_radius_m)
  movel([-0.069296, -0.956555, -2.742713, -1.013120, 1.570796, 1.501500],accel_mss,speed_ms,0,blend_radius_m)
  movel([-0.067994, -0.961593, -2.741336, -1.009460, 1.570796, 1.502802],accel_mss,speed_ms,0,blend_radius_m)
  movel([-0.067482, -0.962340, -2.741130, -1.008919, 1.570796, 1.503314],accel_mss,speed_ms,0,blend_radius_m)
  movel([-0.067015, -0.962322, -2.741135, -1.008932, 1.570796, 1.503782],accel_mss,speed_ms,0,blend_radius_m)
  movel([-0.066333, -0.961956, -2.741236, -1.009197, 1.570796, 1.504463],accel_mss,speed_ms,0,blend_radius_m)
  movel([-0.065449, -0.959415, -2.741934, -1.011041, 1.570796, 1.505347],accel_mss,speed_ms,0,blend_radius_m)
  movel([-0.064723, -0.956867, -2.742629, -1.012893, 1.570796, 1.506074],accel_mss,speed_ms,0,blend_radius_m)
  movel([-0.063159, -0.964473, -2.740540, -1.007376, 1.570796, 1.507637],accel_mss,speed_ms,0,blend_radius_m)
  movel([-0.061322, -0.971801, -2.738489, -1.002099, 1.570796, 1.509475],accel_mss,speed_ms,0,blend_radius_m)
  movel([-0.059217, -0.978853, -2.736479, -0.997057, 1.570796, 1.511580],accel_mss,speed_ms,0,blend_radius_m)
  movel([-0.056851, -0.985636, -2.734510, -0.992243, 1.570796, 1.513946],accel_mss,speed_ms,0,blend_radius_m)
  movel([-0.055705, -0.988480, -2.733675, -0.990234, 1.570796, 1.515091],accel_mss,speed_ms,0,blend_radius_m)
  movel([-0.054214, -0.991193, -2.732873, -0.988323, 1.570796, 1.516582],accel_mss,speed_ms,0,blend_radius_m)
  movel([-0.053288, -0.992366, -2.732524, -0.987499, 1.570796, 1.517508],accel_mss,speed_ms,0,blend_radius_m)
  movel([-0.052214, -0.993345, -2.732232, -0.986812, 1.570796, 1.518582],accel_mss,speed_ms,0,blend_radius_m)
  movel([-0.050968, -0.994073, -2.732015, -0.986301, 1.570796, 1.519828],accel_mss,speed_ms,0,blend_radius_m)
  movel([-0.049530, -0.994493, -2.731889, -0.986007, 1.570796, 1.521266],accel_mss,speed_ms,0,blend_radius_m)
  movel([-0.048410, -0.994565, -2.731868, -0.985957, 1.570796, 1.522386],accel_mss,speed_ms,0,blend_radius_m)
  movel([-0.045989, -0.994112, -2.732003, -0.986274, 1.570796, 1.524807],accel_mss,speed_ms,0,blend_radius_m)
  movel([-0.044708, -0.993619, -2.732150, -0.986620, 1.570796, 1.526088],accel_mss,speed_ms,0,blend_radius_m)
  movel([-0.042057, -0.992185, -2.732578, -0.987626, 1.570796, 1.528740],accel_mss,speed_ms,0,blend_radius_m)
  movel([-0.039350, -0.990250, -2.733152, -0.988987, 1.570796, 1.531447],accel_mss,speed_ms,0,blend_radius_m)
  movel([-0.036671, -0.987945, -2.733833, -0.990611, 1.570796, 1.534126],accel_mss,speed_ms,0,blend_radius_m)
  movel([-0.034103, -0.985390, -2.734582, -0.992416, 1.570796, 1.536693],accel_mss,speed_ms,0,blend_radius_m)
  movel([-0.031730, -0.982718, -2.735361, -0.994309, 1.570796, 1.539066],accel_mss,speed_ms,0,blend_radius_m)
  movel([-0.029646, -0.980059, -2.736131, -0.996199, 1.570796, 1.541150],accel_mss,speed_ms,0,blend_radius_m)
  speed_ms = 0.005
  movel([-0.029646, -0.971223, -2.730367, -1.010798, 1.570796, 1.541150],accel_mss,speed_ms,0,blend_radius_m)
  speed_ms = 0.040
  movel([-0.042131, -0.979992, -2.727833, -1.004565, 1.570796, 1.528666],accel_mss,speed_ms,0,blend_radius_m)
  speed_ms = 0.005
  movel([-0.042131, -0.988862, -2.733563, -0.989965, 1.570796, 1.528666],accel_mss,speed_ms,0,blend_radius_m)
  speed_ms = 0.025
  movel([-0.040484, -0.986656, -2.734212, -0.991522, 1.570796, 1.530312],accel_mss,speed_ms,0,blend_radius_m)
  movel([-0.037383, -0.981853, -2.735612, -0.994923, 1.570796, 1.533413],accel_mss,speed_ms,0,blend_radius_m)
  movel([-0.035957, -0.979308, -2.736348, -0.996733, 1.570796, 1.534839],accel_mss,speed_ms,0,blend_radius_m)
  movel([-0.033421, -0.974060, -2.737849, -1.000480, 1.570796, 1.537375],accel_mss,speed_ms,0,blend_radius_m)
  movel([-0.031384, -0.968766, -2.739343, -1.004280, 1.570796, 1.539412],accel_mss,speed_ms,0,blend_radius_m)
  movel([-0.030589, -0.966172, -2.740068, -1.006149, 1.570796, 1.540208],accel_mss,speed_ms,0,blend_radius_m)
  movel([-0.029964, -0.963646, -2.740769, -1.007974, 1.570796, 1.540833],accel_mss,speed_ms,0,blend_radius_m)
  movel([-0.029275, -0.958922, -2.742069, -1.011399, 1.570796, 1.541522],accel_mss,speed_ms,0,blend_radius_m)
  movel([-0.029237, -0.956774, -2.742654, -1.012961, 1.570796, 1.541560],accel_mss,speed_ms,0,blend_radius_m)
  movel([-0.029428, -0.954816, -2.743185, -1.014388, 1.570796, 1.541368],accel_mss,speed_ms,0,blend_radius_m)
  movel([-0.029858, -0.953070, -2.743656, -1.015663, 1.570796, 1.540939],accel_mss,speed_ms,0,blend_radius_m)
  movel([-0.030542, -0.951566, -2.744060, -1.016763, 1.570796, 1.540254],accel_mss,speed_ms,0,blend_radius_m)
  movel([-0.031674, -0.949978, -2.744485, -1.017925, 1.570796, 1.539122],accel_mss,speed_ms,0,blend_radius_m)
  movel([-0.033044, -0.948663, -2.744836, -1.018890, 1.570796, 1.537752],accel_mss,speed_ms,0,blend_radius_m)
  movel([-0.034661, -0.947691, -2.745094, -1.019603, 1.570796, 1.536136],accel_mss,speed_ms,0,blend_radius_m)
  movel([-0.036529, -0.947136, -2.745242, -1.020012, 1.570796, 1.534267],accel_mss,speed_ms,0,blend_radius_m)
  movel([-0.038659, -0.947065, -2.745260, -1.020063, 1.570796, 1.532137],accel_mss,speed_ms,0,blend_radius_m)
  movel([-0.041047, -0.947550, -2.745132, -1.019708, 1.570796, 1.529749],accel_mss,speed_ms,0,blend_radius_m)
  movel([-0.043700, -0.948658, -2.744837, -1.018894, 1.570796, 1.527096],accel_mss,speed_ms,0,blend_radius_m)
  movel([-0.046618, -0.950447, -2.744360, -1.017582, 1.570796, 1.524178],accel_mss,speed_ms,0,blend_radius_m)
  movel([-0.048590, -0.952011, -2.743941, -1.016437, 1.570796, 1.522206],accel_mss,speed_ms,0,blend_radius_m)
  movel([-0.050473, -0.953828, -2.743452, -1.015109, 1.570796, 1.520324],accel_mss,speed_ms,0,blend_radius_m)
  movel([-0.052203, -0.955822, -2.742913, -1.013655, 1.570796, 1.518593],accel_mss,speed_ms,0,blend_radius_m)
  movel([-0.053730, -0.957924, -2.742341, -1.012124, 1.570796, 1.517066],accel_mss,speed_ms,0,blend_radius_m)
  movel([-0.055002, -0.960067, -2.741755, -1.010567, 1.570796, 1.515794],accel_mss,speed_ms,0,blend_radius_m)
  movel([-0.055966, -0.962182, -2.741174, -1.009034, 1.570796, 1.514831],accel_mss,speed_ms,0,blend_radius_m)
  movel([-0.056566, -0.964199, -2.740616, -1.007574, 1.570796, 1.514231],accel_mss,speed_ms,0,blend_radius_m)
  movel([-0.056759, -0.966058, -2.740100, -1.006231, 1.570796, 1.514037],accel_mss,speed_ms,0,blend_radius_m)
  speed_ms = 0.005
  movel([-0.056759, -0.957281, -2.734283, -1.020824, 1.570796, 1.514037],accel_mss,speed_ms,0,blend_radius_m)
  speed_ms = 0.040
  # Splitting Linear movement in 2 (instruction 399: MoveL 378)
  movel([-0.002283, -0.957501, -2.734223, -1.020666, 1.570796, 1.568514],accel_mss,speed_ms,0,blend_radius_m)
  movel([0.049986, -0.961610, -2.733082, -1.017697, 1.570796, 1.620782],accel_mss,speed_ms,0,blend_radius_m)
  speed_ms = 0.005
  movel([0.049986, -0.970405, -2.738883, -1.003101, 1.570796, 1.620782],accel_mss,speed_ms,0,blend_radius_m)
  speed_ms = 0.025
  movel([0.049190, -0.980201, -2.736090, -0.996098, 1.570796, 1.619986],accel_mss,speed_ms,0,blend_radius_m)
  movel([0.048424, -0.985217, -2.734633, -0.992539, 1.570796, 1.619220],accel_mss,speed_ms,0,blend_radius_m)
  movel([0.047822, -0.987831, -2.733866, -0.990692, 1.570796, 1.618618],accel_mss,speed_ms,0,blend_radius_m)
  movel([0.047025, -0.990539, -2.733067, -0.988783, 1.570796, 1.617821],accel_mss,speed_ms,0,blend_radius_m)
  movel([0.045919, -0.993479, -2.732192, -0.986718, 1.570796, 1.616716],accel_mss,speed_ms,0,blend_radius_m)
  movel([0.045199, -0.994953, -2.731752, -0.985685, 1.570796, 1.615995],accel_mss,speed_ms,0,blend_radius_m)
  movel([0.044310, -0.996412, -2.731314, -0.984664, 1.570796, 1.615106],accel_mss,speed_ms,0,blend_radius_m)
  movel([0.044126, -0.994303, -2.731946, -0.986140, 1.570796, 1.614922],accel_mss,speed_ms,0,blend_radius_m)
  movel([0.043560, -0.992471, -2.732493, -0.987425, 1.570796, 1.614356],accel_mss,speed_ms,0,blend_radius_m)
  movel([0.043149, -0.992049, -2.732619, -0.987722, 1.570796, 1.613945],accel_mss,speed_ms,0,blend_radius_m)
  movel([0.042762, -0.992131, -2.732594, -0.987664, 1.570796, 1.613558],accel_mss,speed_ms,0,blend_radius_m)
  movel([0.042333, -0.992405, -2.732513, -0.987472, 1.570796, 1.613129],accel_mss,speed_ms,0,blend_radius_m)
  movel([0.041502, -0.993266, -2.732256, -0.986867, 1.570796, 1.612298],accel_mss,speed_ms,0,blend_radius_m)
  movel([0.040380, -0.994858, -2.731780, -0.985751, 1.570796, 1.611176],accel_mss,speed_ms,0,blend_radius_m)
  movel([0.039522, -0.996423, -2.731310, -0.984656, 1.570796, 1.610318],accel_mss,speed_ms,0,blend_radius_m)
  movel([0.038878, -0.997962, -2.730846, -0.983580, 1.570796, 1.609674],accel_mss,speed_ms,0,blend_radius_m)
  movel([0.038400, -0.999474, -2.730389, -0.982526, 1.570796, 1.609196],accel_mss,speed_ms,0,blend_radius_m)
  movel([0.037132, -1.005373, -2.728588, -0.978428, 1.570796, 1.607928],accel_mss,speed_ms,0,blend_radius_m)
  movel([0.036202, -1.008880, -2.727505, -0.976004, 1.570796, 1.606999],accel_mss,speed_ms,0,blend_radius_m)
  movel([0.035039, -1.012437, -2.726396, -0.973555, 1.570796, 1.605836],accel_mss,speed_ms,0,blend_radius_m)
  movel([0.033580, -1.016038, -2.725264, -0.971087, 1.570796, 1.604376],accel_mss,speed_ms,0,blend_radius_m)
  movel([0.031763, -1.019655, -2.724117, -0.968617, 1.570796, 1.602559],accel_mss,speed_ms,0,blend_radius_m)
  movel([0.032137, -1.017055, -2.724943, -0.970391, 1.570796, 1.602934],accel_mss,speed_ms,0,blend_radius_m)
  movel([0.031885, -1.014797, -2.725655, -0.971936, 1.570796, 1.602681],accel_mss,speed_ms,0,blend_radius_m)
  movel([0.031682, -1.014325, -2.725804, -0.972260, 1.570796, 1.602478],accel_mss,speed_ms,0,blend_radius_m)
  movel([0.031269, -1.014095, -2.725876, -0.972417, 1.570796, 1.602066],accel_mss,speed_ms,0,blend_radius_m)
  movel([0.030771, -1.014224, -2.725836, -0.972329, 1.570796, 1.601568],accel_mss,speed_ms,0,blend_radius_m)
  movel([0.030229, -1.014588, -2.725721, -0.972080, 1.570796, 1.601025],accel_mss,speed_ms,0,blend_radius_m)
  movel([0.029211, -1.015670, -2.725380, -0.971339, 1.570796, 1.600007],accel_mss,speed_ms,0,blend_radius_m)
  movel([0.028159, -1.017183, -2.724902, -0.970304, 1.570796, 1.598955],accel_mss,speed_ms,0,blend_radius_m)
  movel([0.027287, -1.018733, -2.724410, -0.969246, 1.570796, 1.598083],accel_mss,speed_ms,0,blend_radius_m)
  movel([0.025943, -1.021875, -2.723407, -0.967107, 1.570796, 1.596739],accel_mss,speed_ms,0,blend_radius_m)
  movel([0.023834, -1.028016, -2.721425, -0.962949, 1.570796, 1.594631],accel_mss,speed_ms,0,blend_radius_m)
  movel([0.022396, -1.031463, -2.720298, -0.960628, 1.570796, 1.593192],accel_mss,speed_ms,0,blend_radius_m)
  movel([0.020733, -1.034914, -2.719161, -0.958314, 1.570796, 1.591529],accel_mss,speed_ms,0,blend_radius_m)
  movel([0.018791, -1.038327, -2.718027, -0.956035, 1.570796, 1.589587],accel_mss,speed_ms,0,blend_radius_m)
  movel([0.016519, -1.041664, -2.716909, -0.953816, 1.570796, 1.587315],accel_mss,speed_ms,0,blend_radius_m)
  movel([0.016897, -1.040212, -2.717397, -0.954781, 1.570796, 1.587693],accel_mss,speed_ms,0,blend_radius_m)
  movel([0.017127, -1.037527, -2.718294, -0.956568, 1.570796, 1.587923],accel_mss,speed_ms,0,blend_radius_m)
  movel([0.016973, -1.036334, -2.718691, -0.957365, 1.570796, 1.587769],accel_mss,speed_ms,0,blend_radius_m)
  movel([0.016762, -1.035881, -2.718841, -0.957667, 1.570796, 1.587558],accel_mss,speed_ms,0,blend_radius_m)
  movel([0.016280, -1.035831, -2.718857, -0.957701, 1.570796, 1.587077],accel_mss,speed_ms,0,blend_radius_m)
  movel([0.015644, -1.036371, -2.718678, -0.957340, 1.570796, 1.586440],accel_mss,speed_ms,0,blend_radius_m)
  movel([0.014263, -1.038031, -2.718126, -0.956232, 1.570796, 1.585059],accel_mss,speed_ms,0,blend_radius_m)
  movel([0.013091, -1.039697, -2.717569, -0.955123, 1.570796, 1.583887],accel_mss,speed_ms,0,blend_radius_m)
  movel([0.011129, -1.043052, -2.716441, -0.952895, 1.570796, 1.581925],accel_mss,speed_ms,0,blend_radius_m)
  movel([0.009265, -1.046427, -2.715297, -0.950664, 1.570796, 1.580061],accel_mss,speed_ms,0,blend_radius_m)
  movel([0.008216, -1.048122, -2.714719, -0.949547, 1.570796, 1.579012],accel_mss,speed_ms,0,blend_radius_m)
  movel([0.007006, -1.049824, -2.714137, -0.948429, 1.570796, 1.577802],accel_mss,speed_ms,0,blend_radius_m)
  movel([0.003808, -1.053801, -2.712765, -0.945823, 1.570796, 1.574604],accel_mss,speed_ms,0,blend_radius_m)
  movel([0.000472, -1.057653, -2.711424, -0.943312, 1.570796, 1.571269],accel_mss,speed_ms,0,blend_radius_m)
  movel([-0.002962, -1.061381, -2.710114, -0.940893, 1.570796, 1.567834],accel_mss,speed_ms,0,blend_radius_m)
  movel([-0.006465, -1.065003, -2.708830, -0.938556, 1.570796, 1.564331],accel_mss,speed_ms,0,blend_radius_m)
  speed_ms = 0.005
  movel([-0.006465, -1.055946, -2.703405, -0.953038, 1.570796, 1.564331],accel_mss,speed_ms,0,blend_radius_m)
  speed_ms = 0.040
  movel([-0.038497, -1.032710, -2.711366, -0.968312, 1.570796, 1.532299],accel_mss,speed_ms,0,blend_radius_m)
  speed_ms = 0.005
  movel([-0.038497, -1.041730, -2.716887, -0.953772, 1.570796, 1.532299],accel_mss,speed_ms,0,blend_radius_m)
  speed_ms = 0.025
  movel([-0.037439, -1.040377, -2.717341, -0.954671, 1.570796, 1.533357],accel_mss,speed_ms,0,blend_radius_m)
  movel([-0.036521, -1.038927, -2.717827, -0.955635, 1.570796, 1.534276],accel_mss,speed_ms,0,blend_radius_m)
  movel([-0.034918, -1.035844, -2.718853, -0.957692, 1.570796, 1.535879],accel_mss,speed_ms,0,blend_radius_m)
  movel([-0.033344, -1.032694, -2.719894, -0.959801, 1.570796, 1.537452],accel_mss,speed_ms,0,blend_radius_m)
  movel([-0.032457, -1.031158, -2.720398, -0.960833, 1.570796, 1.538339],accel_mss,speed_ms,0,blend_radius_m)
  movel([-0.031445, -1.029687, -2.720880, -0.961822, 1.570796, 1.539351],accel_mss,speed_ms,0,blend_radius_m)
  movel([-0.030616, -1.028694, -2.721204, -0.962491, 1.570796, 1.540181],accel_mss,speed_ms,0,blend_radius_m)
  movel([-0.029908, -1.028041, -2.721416, -0.962932, 1.570796, 1.540888],accel_mss,speed_ms,0,blend_radius_m)
  movel([-0.029314, -1.027688, -2.721531, -0.963170, 1.570796, 1.541483],accel_mss,speed_ms,0,blend_radius_m)
  movel([-0.028819, -1.027599, -2.721560, -0.963230, 1.570796, 1.541977],accel_mss,speed_ms,0,blend_radius_m)
  movel([-0.028103, -1.028095, -2.721399, -0.962895, 1.570796, 1.542693],accel_mss,speed_ms,0,blend_radius_m)
  movel([-0.027686, -1.029245, -2.721024, -0.962120, 1.570796, 1.543111],accel_mss,speed_ms,0,blend_radius_m)
  movel([-0.027456, -1.032409, -2.719987, -0.959992, 1.570796, 1.543340],accel_mss,speed_ms,0,blend_radius_m)
  movel([-0.027520, -1.034889, -2.719170, -0.958331, 1.570796, 1.543277],accel_mss,speed_ms,0,blend_radius_m)
  movel([-0.025725, -1.031720, -2.720214, -0.960455, 1.570796, 1.545071],accel_mss,speed_ms,0,blend_radius_m)
  movel([-0.024430, -1.028729, -2.721192, -0.962467, 1.570796, 1.546367],accel_mss,speed_ms,0,blend_radius_m)
  movel([-0.023504, -1.025861, -2.722124, -0.964404, 1.570796, 1.547293],accel_mss,speed_ms,0,blend_radius_m)
  movel([-0.022832, -1.023072, -2.723023, -0.966294, 1.570796, 1.547964],accel_mss,speed_ms,0,blend_radius_m)
  movel([-0.021093, -1.014654, -2.725701, -0.972034, 1.570796, 1.549703],accel_mss,speed_ms,0,blend_radius_m)
  movel([-0.020187, -1.011655, -2.726641, -0.974093, 1.570796, 1.550610],accel_mss,speed_ms,0,blend_radius_m)
  movel([-0.019631, -1.010412, -2.727029, -0.974948, 1.570796, 1.551165],accel_mss,speed_ms,0,blend_radius_m)
  movel([-0.019008, -1.009581, -2.727287, -0.975521, 1.570796, 1.551788],accel_mss,speed_ms,0,blend_radius_m)
  movel([-0.018350, -1.009104, -2.727435, -0.975849, 1.570796, 1.552446],accel_mss,speed_ms,0,blend_radius_m)
  movel([-0.017693, -1.008935, -2.727488, -0.975966, 1.570796, 1.553103],accel_mss,speed_ms,0,blend_radius_m)
  movel([-0.017066, -1.009011, -2.727464, -0.975913, 1.570796, 1.553730],accel_mss,speed_ms,0,blend_radius_m)
  movel([-0.016507, -1.009284, -2.727379, -0.975725, 1.570796, 1.554289],accel_mss,speed_ms,0,blend_radius_m)
  movel([-0.015714, -1.010193, -2.727097, -0.975099, 1.570796, 1.555082],accel_mss,speed_ms,0,blend_radius_m)
  movel([-0.015423, -1.011487, -2.726693, -0.974208, 1.570796, 1.555373],accel_mss,speed_ms,0,blend_radius_m)
  movel([-0.015380, -1.013326, -2.726118, -0.972945, 1.570796, 1.555416],accel_mss,speed_ms,0,blend_radius_m)
  movel([-0.015545, -1.016833, -2.725013, -0.970543, 1.570796, 1.555252],accel_mss,speed_ms,0,blend_radius_m)
  movel([-0.013993, -1.010979, -2.726852, -0.974558, 1.570796, 1.556804],accel_mss,speed_ms,0,blend_radius_m)
  movel([-0.013473, -1.008133, -2.727736, -0.976519, 1.570796, 1.557323],accel_mss,speed_ms,0,blend_radius_m)
  movel([-0.012962, -1.002657, -2.729421, -0.980311, 1.570796, 1.557834],accel_mss,speed_ms,0,blend_radius_m)
  movel([-0.012977, -1.000056, -2.730213, -0.982120, 1.570796, 1.557819],accel_mss,speed_ms,0,blend_radius_m)
  movel([-0.013556, -0.995183, -2.731683, -0.985524, 1.570796, 1.557240],accel_mss,speed_ms,0,blend_radius_m)
  speed_ms = 0.005
  movel([-0.013556, -0.986290, -2.725977, -1.000122, 1.570796, 1.557240],accel_mss,speed_ms,0,blend_radius_m)
  speed_ms = 0.040
  movel([-0.030657, -1.012090, -2.718064, -0.982235, 1.570796, 1.540140],accel_mss,speed_ms,0,blend_radius_m)
  speed_ms = 0.005
  movel([-0.030657, -1.021062, -2.723667, -0.967659, 1.570796, 1.540140],accel_mss,speed_ms,0,blend_radius_m)
  speed_ms = 0.025
  movel([-0.032765, -1.024690, -2.722502, -0.965197, 1.570796, 1.538031],accel_mss,speed_ms,0,blend_radius_m)
  movel([-0.034652, -1.028318, -2.721326, -0.962745, 1.570796, 1.536144],accel_mss,speed_ms,0,blend_radius_m)
  movel([-0.038279, -1.035527, -2.718958, -0.957904, 1.570796, 1.532517],accel_mss,speed_ms,0,blend_radius_m)
  movel([-0.040302, -1.039116, -2.717764, -0.955510, 1.570796, 1.530494],accel_mss,speed_ms,0,blend_radius_m)
  movel([-0.042593, -1.042627, -2.716585, -0.953177, 1.570796, 1.528204],accel_mss,speed_ms,0,blend_radius_m)
  movel([-0.045193, -1.045936, -2.715465, -0.950989, 1.570796, 1.525603],accel_mss,speed_ms,0,blend_radius_m)
  movel([-0.046620, -1.047474, -2.714941, -0.949974, 1.570796, 1.524177],accel_mss,speed_ms,0,blend_radius_m)
  movel([-0.048137, -1.048914, -2.714448, -0.949026, 1.570796, 1.522660],accel_mss,speed_ms,0,blend_radius_m)
  movel([-0.047051, -1.047649, -2.714881, -0.949859, 1.570796, 1.523745],accel_mss,speed_ms,0,blend_radius_m)
  movel([-0.045968, -1.045873, -2.715486, -0.951030, 1.570796, 1.524829],accel_mss,speed_ms,0,blend_radius_m)
  movel([-0.045006, -1.043832, -2.716178, -0.952379, 1.570796, 1.525791],accel_mss,speed_ms,0,blend_radius_m)
  movel([-0.044304, -1.041788, -2.716867, -0.953734, 1.570796, 1.526492],accel_mss,speed_ms,0,blend_radius_m)
  movel([-0.043989, -1.039992, -2.717470, -0.954926, 1.570796, 1.526807],accel_mss,speed_ms,0,blend_radius_m)
  movel([-0.044022, -1.039276, -2.717710, -0.955403, 1.570796, 1.526775],accel_mss,speed_ms,0,blend_radius_m)
  movel([-0.044199, -1.038718, -2.717897, -0.955774, 1.570796, 1.526597],accel_mss,speed_ms,0,blend_radius_m)
  movel([-0.044539, -1.038352, -2.718019, -0.956018, 1.570796, 1.526257],accel_mss,speed_ms,0,blend_radius_m)
  movel([-0.045062, -1.038217, -2.718064, -0.956108, 1.570796, 1.525734],accel_mss,speed_ms,0,blend_radius_m)
  movel([-0.045778, -1.038339, -2.718023, -0.956027, 1.570796, 1.525019],accel_mss,speed_ms,0,blend_radius_m)
  movel([-0.046709, -1.038754, -2.717884, -0.955750, 1.570796, 1.524087],accel_mss,speed_ms,0,blend_radius_m)
  movel([-0.048161, -1.039843, -2.717520, -0.955026, 1.570796, 1.522635],accel_mss,speed_ms,0,blend_radius_m)
  movel([-0.053993, -1.045536, -2.715600, -0.951253, 1.570796, 1.516804],accel_mss,speed_ms,0,blend_radius_m)
  movel([-0.056512, -1.047722, -2.714856, -0.949811, 1.570796, 1.514285],accel_mss,speed_ms,0,blend_radius_m)
  movel([-0.059118, -1.049763, -2.714157, -0.948468, 1.570796, 1.511679],accel_mss,speed_ms,0,blend_radius_m)
  movel([-0.061734, -1.051553, -2.713542, -0.947294, 1.570796, 1.509062],accel_mss,speed_ms,0,blend_radius_m)
  movel([-0.064286, -1.052974, -2.713051, -0.946364, 1.570796, 1.506510],accel_mss,speed_ms,0,blend_radius_m)
  movel([-0.066703, -1.053920, -2.712724, -0.945745, 1.570796, 1.504093],accel_mss,speed_ms,0,blend_radius_m)
  movel([-0.068910, -1.054272, -2.712602, -0.945515, 1.570796, 1.501886],accel_mss,speed_ms,0,blend_radius_m)
  movel([-0.068214, -1.054061, -2.712675, -0.945653, 1.570796, 1.502582],accel_mss,speed_ms,0,blend_radius_m)
  movel([-0.067329, -1.053501, -2.712869, -0.946019, 1.570796, 1.503467],accel_mss,speed_ms,0,blend_radius_m)
  movel([-0.065255, -1.051699, -2.713492, -0.947199, 1.570796, 1.505541],accel_mss,speed_ms,0,blend_radius_m)
  movel([-0.063253, -1.049601, -2.714213, -0.948575, 1.570796, 1.507543],accel_mss,speed_ms,0,blend_radius_m)
  movel([-0.061896, -1.047956, -2.714776, -0.949657, 1.570796, 1.508900],accel_mss,speed_ms,0,blend_radius_m)
  movel([-0.061127, -1.046725, -2.715196, -0.950468, 1.570796, 1.509669],accel_mss,speed_ms,0,blend_radius_m)
  movel([-0.060876, -1.045937, -2.715464, -0.950988, 1.570796, 1.509920],accel_mss,speed_ms,0,blend_radius_m)
  movel([-0.061059, -1.045521, -2.715605, -0.951262, 1.570796, 1.509737],accel_mss,speed_ms,0,blend_radius_m)
  movel([-0.061581, -1.045407, -2.715644, -0.951338, 1.570796, 1.509215],accel_mss,speed_ms,0,blend_radius_m)
  movel([-0.063268, -1.045799, -2.715511, -0.951079, 1.570796, 1.507528],accel_mss,speed_ms,0,blend_radius_m)
  movel([-0.065192, -1.046538, -2.715260, -0.950591, 1.570796, 1.505604],accel_mss,speed_ms,0,blend_radius_m)
  movel([-0.069563, -1.048215, -2.714688, -0.949486, 1.570796, 1.501234],accel_mss,speed_ms,0,blend_radius_m)
  movel([-0.073945, -1.049544, -2.714232, -0.948612, 1.570796, 1.496851],accel_mss,speed_ms,0,blend_radius_m)
  movel([-0.076036, -1.049944, -2.714095, -0.948349, 1.570796, 1.494760],accel_mss,speed_ms,0,blend_radius_m)
  movel([-0.078004, -1.050095, -2.714043, -0.948251, 1.570796, 1.492793],accel_mss,speed_ms,0,blend_radius_m)
  movel([-0.079805, -1.049939, -2.714097, -0.948353, 1.570796, 1.490991],accel_mss,speed_ms,0,blend_radius_m)
  movel([-0.081399, -1.049424, -2.714274, -0.948691, 1.570796, 1.489397],accel_mss,speed_ms,0,blend_radius_m)
  movel([-0.078799, -1.048401, -2.714624, -0.949364, 1.570796, 1.491997],accel_mss,speed_ms,0,blend_radius_m)
  movel([-0.077404, -1.047560, -2.714911, -0.949918, 1.570796, 1.493392],accel_mss,speed_ms,0,blend_radius_m)
  movel([-0.076800, -1.047039, -2.715089, -0.950261, 1.570796, 1.493996],accel_mss,speed_ms,0,blend_radius_m)
  movel([-0.076301, -1.046439, -2.715293, -0.950657, 1.570796, 1.494495],accel_mss,speed_ms,0,blend_radius_m)
  movel([-0.076117, -1.046001, -2.715442, -0.950946, 1.570796, 1.494679],accel_mss,speed_ms,0,blend_radius_m)
  movel([-0.076189, -1.045627, -2.715569, -0.951193, 1.570796, 1.494608],accel_mss,speed_ms,0,blend_radius_m)
  movel([-0.076958, -1.045049, -2.715766, -0.951574, 1.570796, 1.493839],accel_mss,speed_ms,0,blend_radius_m)
  movel([-0.078371, -1.044671, -2.715894, -0.951824, 1.570796, 1.492425],accel_mss,speed_ms,0,blend_radius_m)
  movel([-0.080180, -1.044447, -2.715970, -0.951972, 1.570796, 1.490616],accel_mss,speed_ms,0,blend_radius_m)
  movel([-0.086458, -1.044261, -2.716033, -0.952095, 1.570796, 1.484338],accel_mss,speed_ms,0,blend_radius_m)
  movel([-0.088766, -1.043875, -2.716163, -0.952351, 1.570796, 1.482030],accel_mss,speed_ms,0,blend_radius_m)
  movel([-0.090886, -1.043189, -2.716395, -0.952805, 1.570796, 1.479911],accel_mss,speed_ms,0,blend_radius_m)
  movel([-0.092693, -1.042114, -2.716758, -0.953517, 1.570796, 1.478103],accel_mss,speed_ms,0,blend_radius_m)
  movel([-0.094081, -1.040564, -2.717279, -0.954546, 1.570796, 1.476715],accel_mss,speed_ms,0,blend_radius_m)
  movel([-0.091937, -1.041029, -2.717123, -0.954237, 1.570796, 1.478859],accel_mss,speed_ms,0,blend_radius_m)
  movel([-0.090632, -1.041015, -2.717127, -0.954247, 1.570796, 1.480165],accel_mss,speed_ms,0,blend_radius_m)
  movel([-0.089404, -1.040608, -2.717264, -0.954517, 1.570796, 1.481392],accel_mss,speed_ms,0,blend_radius_m)
  movel([-0.088282, -1.039740, -2.717555, -0.955094, 1.570796, 1.482514],accel_mss,speed_ms,0,blend_radius_m)
  movel([-0.087653, -1.038789, -2.717873, -0.955727, 1.570796, 1.483143],accel_mss,speed_ms,0,blend_radius_m)
  movel([-0.087532, -1.037877, -2.718177, -0.956335, 1.570796, 1.483264],accel_mss,speed_ms,0,blend_radius_m)
  movel([-0.087931, -1.037120, -2.718429, -0.956839, 1.570796, 1.482865],accel_mss,speed_ms,0,blend_radius_m)
  movel([-0.090937, -1.033819, -2.719523, -0.959047, 1.570796, 1.479859],accel_mss,speed_ms,0,blend_radius_m)
  movel([-0.093360, -1.030076, -2.720752, -0.961560, 1.570796, 1.477437],accel_mss,speed_ms,0,blend_radius_m)
  movel([-0.094313, -1.027969, -2.721440, -0.962980, 1.570796, 1.476484],accel_mss,speed_ms,0,blend_radius_m)
  movel([-0.095076, -1.025669, -2.722186, -0.964534, 1.570796, 1.475721],accel_mss,speed_ms,0,blend_radius_m)
  movel([-0.095631, -1.023146, -2.722999, -0.966244, 1.570796, 1.475165],accel_mss,speed_ms,0,blend_radius_m)
  movel([-0.095964, -1.020371, -2.723888, -0.968130, 1.570796, 1.474832],accel_mss,speed_ms,0,blend_radius_m)
  speed_ms = 0.005
  movel([-0.095964, -1.011400, -2.718282, -0.982707, 1.570796, 1.474832],accel_mss,speed_ms,0,blend_radius_m)
  speed_ms = 0.040
  movel([-0.138779, -1.008737, -2.719121, -0.984531, 1.570796, 1.432017],accel_mss,speed_ms,0,blend_radius_m)
  speed_ms = 0.005
  movel([-0.138779, -1.017700, -2.724738, -0.969950, 1.570796, 1.432017],accel_mss,speed_ms,0,blend_radius_m)
  speed_ms = 0.025
  movel([-0.135945, -1.012396, -2.726409, -0.973584, 1.570796, 1.434851],accel_mss,speed_ms,0,blend_radius_m)
  movel([-0.133243, -1.007057, -2.728069, -0.977263, 1.570796, 1.437553],accel_mss,speed_ms,0,blend_radius_m)
  movel([-0.128172, -0.996240, -2.731365, -0.984784, 1.570796, 1.442625],accel_mss,speed_ms,0,blend_radius_m)
  movel([-0.123556, -0.985275, -2.734616, -0.992498, 1.570796, 1.447241],accel_mss,speed_ms,0,blend_radius_m)
  movel([-0.119410, -0.974201, -2.737809, -1.000379, 1.570796, 1.451386],accel_mss,speed_ms,0,blend_radius_m)
  movel([-0.115748, -0.963054, -2.740933, -1.008402, 1.570796, 1.455048],accel_mss,speed_ms,0,blend_radius_m)
  movel([-0.112588, -0.951883, -2.743975, -1.016531, 1.570796, 1.458208],accel_mss,speed_ms,0,blend_radius_m)
  movel([-0.109947, -0.940739, -2.746924, -1.024727, 1.570796, 1.460850],accel_mss,speed_ms,0,blend_radius_m)
  movel([-0.107841, -0.929667, -2.749769, -1.032953, 1.570796, 1.462955],accel_mss,speed_ms,0,blend_radius_m)
  movel([-0.106293, -0.918734, -2.752499, -1.041157, 1.570796, 1.464503],accel_mss,speed_ms,0,blend_radius_m)
  movel([-0.105324, -0.907996, -2.755103, -1.049290, 1.570796, 1.465473],accel_mss,speed_ms,0,blend_radius_m)
  movel([-0.104957, -0.897520, -2.757573, -1.057296, 1.570796, 1.465840],accel_mss,speed_ms,0,blend_radius_m)
  movel([-0.105217, -0.887377, -2.759898, -1.065114, 1.570796, 1.465579],accel_mss,speed_ms,0,blend_radius_m)
  movel([-0.106118, -0.877626, -2.762073, -1.072690, 1.570796, 1.464678],accel_mss,speed_ms,0,blend_radius_m)
  movel([-0.107693, -0.868355, -2.764088, -1.079946, 1.570796, 1.463104],accel_mss,speed_ms,0,blend_radius_m)
  movel([-0.109956, -0.859634, -2.765936, -1.086819, 1.570796, 1.460840],accel_mss,speed_ms,0,blend_radius_m)
  movel([-0.114456, -0.847511, -2.768431, -1.096447, 1.570796, 1.456341],accel_mss,speed_ms,0,blend_radius_m)
  movel([-0.114855, -0.845201, -2.768896, -1.098292, 1.570796, 1.455941],accel_mss,speed_ms,0,blend_radius_m)
  movel([-0.114786, -0.842543, -2.769429, -1.100418, 1.570796, 1.456010],accel_mss,speed_ms,0,blend_radius_m)
  movel([-0.114004, -0.838474, -2.770235, -1.103679, 1.570796, 1.456792],accel_mss,speed_ms,0,blend_radius_m)
  movel([-0.112787, -0.835025, -2.770911, -1.106452, 1.570796, 1.458009],accel_mss,speed_ms,0,blend_radius_m)
  movel([-0.112035, -0.833525, -2.771204, -1.107660, 1.570796, 1.458762],accel_mss,speed_ms,0,blend_radius_m)
  movel([-0.110274, -0.830935, -2.771705, -1.109749, 1.570796, 1.460522],accel_mss,speed_ms,0,blend_radius_m)
  movel([-0.109287, -0.829846, -2.771915, -1.110629, 1.570796, 1.461509],accel_mss,speed_ms,0,blend_radius_m)
  movel([-0.107116, -0.828036, -2.772262, -1.112091, 1.570796, 1.463681],accel_mss,speed_ms,0,blend_radius_m)
  movel([-0.104747, -0.826695, -2.772518, -1.113176, 1.570796, 1.466049],accel_mss,speed_ms,0,blend_radius_m)
  movel([-0.102241, -0.825783, -2.772691, -1.113915, 1.570796, 1.468556],accel_mss,speed_ms,0,blend_radius_m)
  movel([-0.099652, -0.825259, -2.772791, -1.114339, 1.570796, 1.471145],accel_mss,speed_ms,0,blend_radius_m)
  movel([-0.097045, -0.825078, -2.772825, -1.114486, 1.570796, 1.473752],accel_mss,speed_ms,0,blend_radius_m)
  movel([-0.094473, -0.825200, -2.772802, -1.114387, 1.570796, 1.476323],accel_mss,speed_ms,0,blend_radius_m)
  movel([-0.089682, -0.826157, -2.772620, -1.113612, 1.570796, 1.481114],accel_mss,speed_ms,0,blend_radius_m)
  movel([-0.085723, -0.827757, -2.772315, -1.112317, 1.570796, 1.485073],accel_mss,speed_ms,0,blend_radius_m)
  movel([-0.083017, -0.829586, -2.771965, -1.110839, 1.570796, 1.487779],accel_mss,speed_ms,0,blend_radius_m)
  movel([-0.080464, -0.832402, -2.771421, -1.108565, 1.570796, 1.490333],accel_mss,speed_ms,0,blend_radius_m)
  movel([-0.078266, -0.835611, -2.770797, -1.105981, 1.570796, 1.492531],accel_mss,speed_ms,0,blend_radius_m)
  movel([-0.074605, -0.842784, -2.769380, -1.100225, 1.570796, 1.496191],accel_mss,speed_ms,0,blend_radius_m)
  movel([-0.071379, -0.850312, -2.767862, -1.094215, 1.570796, 1.499418],accel_mss,speed_ms,0,blend_radius_m)
  movel([-0.067955, -0.857444, -2.766393, -1.088552, 1.570796, 1.502841],accel_mss,speed_ms,0,blend_radius_m)
  movel([-0.064391, -0.863299, -2.765165, -1.083925, 1.570796, 1.506406],accel_mss,speed_ms,0,blend_radius_m)
  movel([-0.062241, -0.865799, -2.764634, -1.081956, 1.570796, 1.508556],accel_mss,speed_ms,0,blend_radius_m)
  movel([-0.059643, -0.867756, -2.764216, -1.080417, 1.570796, 1.511154],accel_mss,speed_ms,0,blend_radius_m)
  movel([-0.058167, -0.868326, -2.764094, -1.079969, 1.570796, 1.512630],accel_mss,speed_ms,0,blend_radius_m)
  movel([-0.057282, -0.868359, -2.764087, -1.079943, 1.570796, 1.513515],accel_mss,speed_ms,0,blend_radius_m)
  movel([-0.056273, -0.868126, -2.764137, -1.080126, 1.570796, 1.514524],accel_mss,speed_ms,0,blend_radius_m)
  movel([-0.054860, -0.867396, -2.764293, -1.080700, 1.570796, 1.515936],accel_mss,speed_ms,0,blend_radius_m)
  movel([-0.053419, -0.866298, -2.764528, -1.081563, 1.570796, 1.517377],accel_mss,speed_ms,0,blend_radius_m)
  movel([-0.050618, -0.863492, -2.765124, -1.083773, 1.570796, 1.520178],accel_mss,speed_ms,0,blend_radius_m)
  movel([-0.047614, -0.859986, -2.765862, -1.086541, 1.570796, 1.523182],accel_mss,speed_ms,0,blend_radius_m)
  movel([-0.044782, -0.856365, -2.766617, -1.089407, 1.570796, 1.526014],accel_mss,speed_ms,0,blend_radius_m)
  movel([-0.039495, -0.848855, -2.768158, -1.095376, 1.570796, 1.531301],accel_mss,speed_ms,0,blend_radius_m)
  movel([-0.029331, -0.833325, -2.771242, -1.107821, 1.570796, 1.541466],accel_mss,speed_ms,0,blend_radius_m)
  movel([-0.024263, -0.826028, -2.772645, -1.113716, 1.570796, 1.546533],accel_mss,speed_ms,0,blend_radius_m)
  movel([-0.021239, -0.822033, -2.773400, -1.116956, 1.570796, 1.549558],accel_mss,speed_ms,0,blend_radius_m)
  movel([-0.018125, -0.818369, -2.774084, -1.119936, 1.570796, 1.552671],accel_mss,speed_ms,0,blend_radius_m)
  movel([-0.016592, -0.816790, -2.774377, -1.121221, 1.570796, 1.554204],accel_mss,speed_ms,0,blend_radius_m)
  movel([-0.015103, -0.815453, -2.774624, -1.122312, 1.570796, 1.555693],accel_mss,speed_ms,0,blend_radius_m)
  movel([-0.013687, -0.814411, -2.774816, -1.123162, 1.570796, 1.557109],accel_mss,speed_ms,0,blend_radius_m)
  movel([-0.012363, -0.813721, -2.774942, -1.123726, 1.570796, 1.558433],accel_mss,speed_ms,0,blend_radius_m)
  movel([-0.011160, -0.813431, -2.774995, -1.123962, 1.570796, 1.559636],accel_mss,speed_ms,0,blend_radius_m)
  movel([-0.010099, -0.813595, -2.774966, -1.123829, 1.570796, 1.560697],accel_mss,speed_ms,0,blend_radius_m)
  movel([-0.009203, -0.814268, -2.774842, -1.123279, 1.570796, 1.561593],accel_mss,speed_ms,0,blend_radius_m)
  movel([-0.008500, -0.815504, -2.774615, -1.122270, 1.570796, 1.562296],accel_mss,speed_ms,0,blend_radius_m)
  movel([-0.007699, -0.818093, -2.774136, -1.120161, 1.570796, 1.563097],accel_mss,speed_ms,0,blend_radius_m)
  movel([-0.007237, -0.820886, -2.773615, -1.117888, 1.570796, 1.563559],accel_mss,speed_ms,0,blend_radius_m)
  movel([-0.007092, -0.823859, -2.773056, -1.115474, 1.570796, 1.563704],accel_mss,speed_ms,0,blend_radius_m)
  movel([-0.007242, -0.826998, -2.772460, -1.112931, 1.570796, 1.563554],accel_mss,speed_ms,0,blend_radius_m)
  movel([-0.007676, -0.830277, -2.771832, -1.110280, 1.570796, 1.563120],accel_mss,speed_ms,0,blend_radius_m)
  movel([-0.008372, -0.833681, -2.771173, -1.107535, 1.570796, 1.562425],accel_mss,speed_ms,0,blend_radius_m)
  movel([-0.009313, -0.837192, -2.770487, -1.104710, 1.570796, 1.561483],accel_mss,speed_ms,0,blend_radius_m)
  movel([-0.010479, -0.840792, -2.769777, -1.101820, 1.570796, 1.560317],accel_mss,speed_ms,0,blend_radius_m)
  movel([-0.013418, -0.848180, -2.768295, -1.095914, 1.570796, 1.557379],accel_mss,speed_ms,0,blend_radius_m)
  movel([-0.017054, -0.855721, -2.766751, -1.089918, 1.570796, 1.553742],accel_mss,speed_ms,0,blend_radius_m)
  movel([-0.021261, -0.863287, -2.765167, -1.083935, 1.570796, 1.549535],accel_mss,speed_ms,0,blend_radius_m)
  movel([-0.025902, -0.870754, -2.763571, -1.078063, 1.570796, 1.544894],accel_mss,speed_ms,0,blend_radius_m)
  movel([-0.036656, -0.887094, -2.759962, -1.065333, 1.570796, 1.534140],accel_mss,speed_ms,0,blend_radius_m)
  movel([-0.042378, -0.895077, -2.758138, -1.059173, 1.570796, 1.528418],accel_mss,speed_ms,0,blend_radius_m)
  movel([-0.045329, -0.898848, -2.757264, -1.056278, 1.570796, 1.525467],accel_mss,speed_ms,0,blend_radius_m)
  movel([-0.048348, -0.902409, -2.756429, -1.053551, 1.570796, 1.522449],accel_mss,speed_ms,0,blend_radius_m)
  movel([-0.050333, -0.904549, -2.755923, -1.051917, 1.570796, 1.520464],accel_mss,speed_ms,0,blend_radius_m)
  movel([-0.052344, -0.906507, -2.755458, -1.050424, 1.570796, 1.518452],accel_mss,speed_ms,0,blend_radius_m)
  movel([-0.054371, -0.908254, -2.755041, -1.049094, 1.570796, 1.516425],accel_mss,speed_ms,0,blend_radius_m)
  movel([-0.056400, -0.909759, -2.754681, -1.047950, 1.570796, 1.514396],accel_mss,speed_ms,0,blend_radius_m)
  movel([-0.058414, -0.910992, -2.754384, -1.047013, 1.570796, 1.512383],accel_mss,speed_ms,0,blend_radius_m)
  movel([-0.060402, -0.911925, -2.754159, -1.046306, 1.570796, 1.510394],accel_mss,speed_ms,0,blend_radius_m)
  movel([-0.062348, -0.912520, -2.754015, -1.045855, 1.570796, 1.508448],accel_mss,speed_ms,0,blend_radius_m)
  movel([-0.064243, -0.912748, -2.753960, -1.045681, 1.570796, 1.506553],accel_mss,speed_ms,0,blend_radius_m)
  movel([-0.066004, -0.912571, -2.754003, -1.045816, 1.570796, 1.504792],accel_mss,speed_ms,0,blend_radius_m)
  movel([-0.067515, -0.912048, -2.754129, -1.046212, 1.570796, 1.503281],accel_mss,speed_ms,0,blend_radius_m)
  movel([-0.072772, -0.908794, -2.754912, -1.048683, 1.570796, 1.498024],accel_mss,speed_ms,0,blend_radius_m)
  movel([-0.074325, -0.908270, -2.755037, -1.049081, 1.570796, 1.496472],accel_mss,speed_ms,0,blend_radius_m)
  movel([-0.076147, -0.908102, -2.755078, -1.049210, 1.570796, 1.494649],accel_mss,speed_ms,0,blend_radius_m)
  movel([-0.076946, -0.908287, -2.755033, -1.049068, 1.570796, 1.493850],accel_mss,speed_ms,0,blend_radius_m)
  movel([-0.077268, -0.908768, -2.754918, -1.048703, 1.570796, 1.493528],accel_mss,speed_ms,0,blend_radius_m)
  movel([-0.077634, -0.909826, -2.754664, -1.047898, 1.570796, 1.493162],accel_mss,speed_ms,0,blend_radius_m)
  movel([-0.078488, -0.913377, -2.753807, -1.045205, 1.570796, 1.492309],accel_mss,speed_ms,0,blend_radius_m)
  movel([-0.080403, -0.923906, -2.751217, -1.037266, 1.570796, 1.490393],accel_mss,speed_ms,0,blend_radius_m)
  movel([-0.083269, -0.941281, -2.746782, -1.024326, 1.570796, 1.487527],accel_mss,speed_ms,0,blend_radius_m)
  movel([-0.085739, -0.950710, -2.744290, -1.017390, 1.570796, 1.485058],accel_mss,speed_ms,0,blend_radius_m)
  movel([-0.088602, -0.960170, -2.741727, -1.010492, 1.570796, 1.482194],accel_mss,speed_ms,0,blend_radius_m)
  movel([-0.091810, -0.969628, -2.739101, -1.003660, 1.570796, 1.478986],accel_mss,speed_ms,0,blend_radius_m)
  movel([-0.095299, -0.979038, -2.736425, -0.996926, 1.570796, 1.475497],accel_mss,speed_ms,0,blend_radius_m)
  movel([-0.099991, -0.990981, -2.732936, -0.988472, 1.570796, 1.470805],accel_mss,speed_ms,0,blend_radius_m)
  movel([-0.104876, -1.002822, -2.729370, -0.980197, 1.570796, 1.465920],accel_mss,speed_ms,0,blend_radius_m)
  movel([-0.110005, -1.014521, -2.725742, -0.972126, 1.570796, 1.460791],accel_mss,speed_ms,0,blend_radius_m)
  movel([-0.115440, -1.026044, -2.722065, -0.964281, 1.570796, 1.455357],accel_mss,speed_ms,0,blend_radius_m)
  movel([-0.121230, -1.037348, -2.718353, -0.956687, 1.570796, 1.449566],accel_mss,speed_ms,0,blend_radius_m)
  movel([-0.124272, -1.042908, -2.716490, -0.952991, 1.570796, 1.446524],accel_mss,speed_ms,0,blend_radius_m)
  movel([-0.127426, -1.048405, -2.714623, -0.949361, 1.570796, 1.443371],accel_mss,speed_ms,0,blend_radius_m)
  movel([-0.130696, -1.053834, -2.712754, -0.945801, 1.570796, 1.440101],accel_mss,speed_ms,0,blend_radius_m)
  movel([-0.134086, -1.059187, -2.710887, -0.942315, 1.570796, 1.436710],accel_mss,speed_ms,0,blend_radius_m)
  movel([-0.137604, -1.064468, -2.709021, -0.938900, 1.570796, 1.433192],accel_mss,speed_ms,0,blend_radius_m)
  movel([-0.141261, -1.069668, -2.707160, -0.935561, 1.570796, 1.429535],accel_mss,speed_ms,0,blend_radius_m)
  movel([-0.145763, -1.075734, -2.704960, -0.931695, 1.570796, 1.425033],accel_mss,speed_ms,0,blend_radius_m)
  movel([-0.148132, -1.078666, -2.703885, -0.929838, 1.570796, 1.422664],accel_mss,speed_ms,0,blend_radius_m)
  movel([-0.152454, -1.083423, -2.702125, -0.926841, 1.570796, 1.418343],accel_mss,speed_ms,0,blend_radius_m)
  movel([-0.154719, -1.085620, -2.701305, -0.925464, 1.570796, 1.416078],accel_mss,speed_ms,0,blend_radius_m)
  movel([-0.157041, -1.087421, -2.700630, -0.924338, 1.570796, 1.413756],accel_mss,speed_ms,0,blend_radius_m)
  movel([-0.158104, -1.087970, -2.700424, -0.923995, 1.570796, 1.412692],accel_mss,speed_ms,0,blend_radius_m)
  movel([-0.159046, -1.088181, -2.700344, -0.923864, 1.570796, 1.411751],accel_mss,speed_ms,0,blend_radius_m)
  movel([-0.158634, -1.085765, -2.701251, -0.925373, 1.570796, 1.412162],accel_mss,speed_ms,0,blend_radius_m)
  movel([-0.158574, -1.083507, -2.702094, -0.926789, 1.570796, 1.412222],accel_mss,speed_ms,0,blend_radius_m)
  movel([-0.158757, -1.082551, -2.702449, -0.927389, 1.570796, 1.412040],accel_mss,speed_ms,0,blend_radius_m)
  movel([-0.159125, -1.081774, -2.702738, -0.927878, 1.570796, 1.411672],accel_mss,speed_ms,0,blend_radius_m)
  movel([-0.159709, -1.081217, -2.702944, -0.928228, 1.570796, 1.411087],accel_mss,speed_ms,0,blend_radius_m)
  movel([-0.160549, -1.080937, -2.703047, -0.928405, 1.570796, 1.410247],accel_mss,speed_ms,0,blend_radius_m)
  movel([-0.163030, -1.080952, -2.703042, -0.928395, 1.570796, 1.407766],accel_mss,speed_ms,0,blend_radius_m)
  movel([-0.163747, -1.080703, -2.703134, -0.928552, 1.570796, 1.407049],accel_mss,speed_ms,0,blend_radius_m)
  movel([-0.164276, -1.080240, -2.703305, -0.928844, 1.570796, 1.406521],accel_mss,speed_ms,0,blend_radius_m)
  movel([-0.164838, -1.078808, -2.703833, -0.929748, 1.570796, 1.405959],accel_mss,speed_ms,0,blend_radius_m)
  movel([-0.164910, -1.076935, -2.704521, -0.930933, 1.570796, 1.405886],accel_mss,speed_ms,0,blend_radius_m)
  movel([-0.164678, -1.074901, -2.705264, -0.932224, 1.570796, 1.406119],accel_mss,speed_ms,0,blend_radius_m)
  movel([-0.163569, -1.068603, -2.707543, -0.936243, 1.570796, 1.407228],accel_mss,speed_ms,0,blend_radius_m)
  movel([-0.162067, -1.062066, -2.709872, -0.940451, 1.570796, 1.408729],accel_mss,speed_ms,0,blend_radius_m)
  movel([-0.161097, -1.058716, -2.711052, -0.942621, 1.570796, 1.409699],accel_mss,speed_ms,0,blend_radius_m)
  movel([-0.159947, -1.055313, -2.712240, -0.944836, 1.570796, 1.410849],accel_mss,speed_ms,0,blend_radius_m)
  movel([-0.158586, -1.051863, -2.713435, -0.947091, 1.570796, 1.412211],accel_mss,speed_ms,0,blend_radius_m)
  movel([-0.156983, -1.048365, -2.714636, -0.949387, 1.570796, 1.413814],accel_mss,speed_ms,0,blend_radius_m)
  movel([-0.155089, -1.044956, -2.715797, -0.951636, 1.570796, 1.415707],accel_mss,speed_ms,0,blend_radius_m)
  movel([-0.148559, -1.035008, -2.719130, -0.958251, 1.570796, 1.422238],accel_mss,speed_ms,0,blend_radius_m)
  movel([-0.143588, -1.026433, -2.721939, -0.964018, 1.570796, 1.427208],accel_mss,speed_ms,0,blend_radius_m)
  movel([-0.138779, -1.017700, -2.724738, -0.969950, 1.570796, 1.432017],accel_mss,speed_ms,0,blend_radius_m)
  movel([-0.136660, -1.013730, -2.725991, -0.972668, 1.570796, 1.434136],accel_mss,speed_ms,0,blend_radius_m)
  speed_ms = 0.005
  movel([-0.136660, -1.004778, -2.720358, -0.987253, 1.570796, 1.434136],accel_mss,speed_ms,0,blend_radius_m)
  speed_ms = 0.040
  movel([-0.181287, -1.075881, -2.696211, -0.940297, 1.570796, 1.389509],accel_mss,speed_ms,0,blend_radius_m)
  speed_ms = 0.005
  movel([-0.181287, -1.084956, -2.701554, -0.925880, 1.570796, 1.389509],accel_mss,speed_ms,0,blend_radius_m)
  speed_ms = 0.025
  movel([-0.176470, -1.087312, -2.700671, -0.924406, 1.570796, 1.394326],accel_mss,speed_ms,0,blend_radius_m)
  movel([-0.174061, -1.088766, -2.700124, -0.923499, 1.570796, 1.396736],accel_mss,speed_ms,0,blend_radius_m)
  movel([-0.171818, -1.090458, -2.699485, -0.922446, 1.570796, 1.398978],accel_mss,speed_ms,0,blend_radius_m)
  movel([-0.169856, -1.092412, -2.698744, -0.921233, 1.570796, 1.400940],accel_mss,speed_ms,0,blend_radius_m)
  movel([-0.168298, -1.094657, -2.697888, -0.919844, 1.570796, 1.402498],accel_mss,speed_ms,0,blend_radius_m)
  movel([-0.167259, -1.097226, -2.696903, -0.918260, 1.570796, 1.403538],accel_mss,speed_ms,0,blend_radius_m)
  movel([-0.166971, -1.098642, -2.696358, -0.917389, 1.570796, 1.403825],accel_mss,speed_ms,0,blend_radius_m)
  movel([-0.166857, -1.100144, -2.695777, -0.916468, 1.570796, 1.403940],accel_mss,speed_ms,0,blend_radius_m)
  movel([-0.167979, -1.099958, -2.695849, -0.916582, 1.570796, 1.402817],accel_mss,speed_ms,0,blend_radius_m)
  movel([-0.168748, -1.099486, -2.696032, -0.916871, 1.570796, 1.402048],accel_mss,speed_ms,0,blend_radius_m)
  movel([-0.170388, -1.098335, -2.696476, -0.917578, 1.570796, 1.400409],accel_mss,speed_ms,0,blend_radius_m)
  movel([-0.172549, -1.097606, -2.696757, -0.918026, 1.570796, 1.398247],accel_mss,speed_ms,0,blend_radius_m)
  movel([-0.174897, -1.097148, -2.696933, -0.918308, 1.570796, 1.395899],accel_mss,speed_ms,0,blend_radius_m)
  movel([-0.177407, -1.096945, -2.697011, -0.918433, 1.570796, 1.393390],accel_mss,speed_ms,0,blend_radius_m)
  movel([-0.180052, -1.096990, -2.696994, -0.918405, 1.570796, 1.390744],accel_mss,speed_ms,0,blend_radius_m)
  movel([-0.182808, -1.097270, -2.696886, -0.918233, 1.570796, 1.387989],accel_mss,speed_ms,0,blend_radius_m)
  movel([-0.185646, -1.097776, -2.696691, -0.917921, 1.570796, 1.385150],accel_mss,speed_ms,0,blend_radius_m)
  movel([-0.188544, -1.098499, -2.696413, -0.917477, 1.570796, 1.382252],accel_mss,speed_ms,0,blend_radius_m)
  movel([-0.191473, -1.099421, -2.696057, -0.916911, 1.570796, 1.379323],accel_mss,speed_ms,0,blend_radius_m)
  movel([-0.193430, -1.100190, -2.695759, -0.916440, 1.570796, 1.377366],accel_mss,speed_ms,0,blend_radius_m)
  movel([-0.194957, -1.100979, -2.695453, -0.915956, 1.570796, 1.375840],accel_mss,speed_ms,0,blend_radius_m)
  movel([-0.196085, -1.101779, -2.695143, -0.915467, 1.570796, 1.374712],accel_mss,speed_ms,0,blend_radius_m)
  movel([-0.196852, -1.102583, -2.694830, -0.914976, 1.570796, 1.373945],accel_mss,speed_ms,0,blend_radius_m)
  movel([-0.197296, -1.103394, -2.694514, -0.914481, 1.570796, 1.373500],accel_mss,speed_ms,0,blend_radius_m)
  movel([-0.197451, -1.104204, -2.694198, -0.913988, 1.570796, 1.373345],accel_mss,speed_ms,0,blend_radius_m)
  movel([-0.197361, -1.105012, -2.693881, -0.913496, 1.570796, 1.373435],accel_mss,speed_ms,0,blend_radius_m)
  movel([-0.197056, -1.105813, -2.693567, -0.913009, 1.570796, 1.373740],accel_mss,speed_ms,0,blend_radius_m)
  movel([-0.195961, -1.107387, -2.692948, -0.912053, 1.570796, 1.374835],accel_mss,speed_ms,0,blend_radius_m)
  movel([-0.191406, -1.111684, -2.691247, -0.909457, 1.570796, 1.379390],accel_mss,speed_ms,0,blend_radius_m)
  movel([-0.194138, -1.111085, -2.691485, -0.909818, 1.570796, 1.376659],accel_mss,speed_ms,0,blend_radius_m)
  movel([-0.199505, -1.109762, -2.692010, -0.910616, 1.570796, 1.371291],accel_mss,speed_ms,0,blend_radius_m)
  movel([-0.202461, -1.109570, -2.692086, -0.910733, 1.570796, 1.368335],accel_mss,speed_ms,0,blend_radius_m)
  movel([-0.205956, -1.109812, -2.691991, -0.910587, 1.570796, 1.364840],accel_mss,speed_ms,0,blend_radius_m)
  movel([-0.209553, -1.110256, -2.691815, -0.910319, 1.570796, 1.361243],accel_mss,speed_ms,0,blend_radius_m)
  movel([-0.216810, -1.111306, -2.691398, -0.909686, 1.570796, 1.353986],accel_mss,speed_ms,0,blend_radius_m)
  movel([-0.220352, -1.111691, -2.691245, -0.909454, 1.570796, 1.350444],accel_mss,speed_ms,0,blend_radius_m)
  movel([-0.223757, -1.111835, -2.691187, -0.909367, 1.570796, 1.347040],accel_mss,speed_ms,0,blend_radius_m)
  movel([-0.226966, -1.111633, -2.691268, -0.909488, 1.570796, 1.343830],accel_mss,speed_ms,0,blend_radius_m)
  movel([-0.229926, -1.110969, -2.691531, -0.909888, 1.570796, 1.340870],accel_mss,speed_ms,0,blend_radius_m)
  movel([-0.226646, -1.114823, -2.689994, -0.907573, 1.570796, 1.344150],accel_mss,speed_ms,0,blend_radius_m)
  movel([-0.224823, -1.116665, -2.689254, -0.906470, 1.570796, 1.345973],accel_mss,speed_ms,0,blend_radius_m)
  movel([-0.222856, -1.118079, -2.688683, -0.905627, 1.570796, 1.347941],accel_mss,speed_ms,0,blend_radius_m)
  movel([-0.225826, -1.117529, -2.688905, -0.905954, 1.570796, 1.344970],accel_mss,speed_ms,0,blend_radius_m)
  movel([-0.229007, -1.117339, -2.688982, -0.906068, 1.570796, 1.341789],accel_mss,speed_ms,0,blend_radius_m)
  movel([-0.235578, -1.117324, -2.688988, -0.906077, 1.570796, 1.335219],accel_mss,speed_ms,0,blend_radius_m)
  movel([-0.237686, -1.117148, -2.689059, -0.906182, 1.570796, 1.333111],accel_mss,speed_ms,0,blend_radius_m)
  movel([-0.239603, -1.116751, -2.689219, -0.906419, 1.570796, 1.331193],accel_mss,speed_ms,0,blend_radius_m)
  movel([-0.243071, -1.115514, -2.689717, -0.907159, 1.570796, 1.327725],accel_mss,speed_ms,0,blend_radius_m)
  movel([-0.246411, -1.114075, -2.690293, -0.908021, 1.570796, 1.324385],accel_mss,speed_ms,0,blend_radius_m)
  movel([-0.250050, -1.112909, -2.690759, -0.908721, 1.570796, 1.320746],accel_mss,speed_ms,0,blend_radius_m)
  movel([-0.251314, -1.112715, -2.690837, -0.908838, 1.570796, 1.319482],accel_mss,speed_ms,0,blend_radius_m)
  movel([-0.252695, -1.112742, -2.690826, -0.908821, 1.570796, 1.318101],accel_mss,speed_ms,0,blend_radius_m)
  movel([-0.254154, -1.113125, -2.690673, -0.908591, 1.570796, 1.316643],accel_mss,speed_ms,0,blend_radius_m)
  movel([-0.254894, -1.113485, -2.690529, -0.908375, 1.570796, 1.315902],accel_mss,speed_ms,0,blend_radius_m)
  movel([-0.255638, -1.113984, -2.690330, -0.908075, 1.570796, 1.315158],accel_mss,speed_ms,0,blend_radius_m)
  movel([-0.256406, -1.114660, -2.690059, -0.907670, 1.570796, 1.314391],accel_mss,speed_ms,0,blend_radius_m)
  movel([-0.257064, -1.115413, -2.689757, -0.907219, 1.570796, 1.313732],accel_mss,speed_ms,0,blend_radius_m)
  movel([-0.258107, -1.117085, -2.689085, -0.906220, 1.570796, 1.312689],accel_mss,speed_ms,0,blend_radius_m)
  movel([-0.258843, -1.118857, -2.688369, -0.905163, 1.570796, 1.311953],accel_mss,speed_ms,0,blend_radius_m)
  movel([-0.259348, -1.120587, -2.687667, -0.904135, 1.570796, 1.311449],accel_mss,speed_ms,0,blend_radius_m)
  movel([-0.260633, -1.118620, -2.688465, -0.905304, 1.570796, 1.310163],accel_mss,speed_ms,0,blend_radius_m)
  movel([-0.262121, -1.116891, -2.689163, -0.906335, 1.570796, 1.308675],accel_mss,speed_ms,0,blend_radius_m)
  movel([-0.265486, -1.113905, -2.690361, -0.908123, 1.570796, 1.305311],accel_mss,speed_ms,0,blend_radius_m)
  movel([-0.269008, -1.111101, -2.691479, -0.909809, 1.570796, 1.301789],accel_mss,speed_ms,0,blend_radius_m)
  movel([-0.272248, -1.107933, -2.692733, -0.911723, 1.570796, 1.298548],accel_mss,speed_ms,0,blend_radius_m)
  movel([-0.273243, -1.106445, -2.693319, -0.912625, 1.570796, 1.297553],accel_mss,speed_ms,0,blend_radius_m)
  movel([-0.273996, -1.104691, -2.694007, -0.913691, 1.570796, 1.296800],accel_mss,speed_ms,0,blend_radius_m)
  movel([-0.274539, -1.102720, -2.694776, -0.914892, 1.570796, 1.296257],accel_mss,speed_ms,0,blend_radius_m)
  movel([-0.274907, -1.100594, -2.695603, -0.916192, 1.570796, 1.295889],accel_mss,speed_ms,0,blend_radius_m)
  movel([-0.275228, -1.096062, -2.697350, -0.918977, 1.570796, 1.295568],accel_mss,speed_ms,0,blend_radius_m)
  movel([-0.275212, -1.091534, -2.699077, -0.921778, 1.570796, 1.295584],accel_mss,speed_ms,0,blend_radius_m)
  speed_ms = 0.005
  movel([-0.275212, -1.082457, -2.693762, -0.936170, 1.570796, 1.295584],accel_mss,speed_ms,0,blend_radius_m)
  speed_ms = 0.040
  # Splitting Linear movement in 2 (instruction 806: MoveL 765)
  movel([-0.254640, -1.013628, -2.717576, -0.981185, 1.570796, 1.316156],accel_mss,speed_ms,0,blend_radius_m)
  movel([-0.230779, -0.937262, -2.739666, -1.035461, 1.570796, 1.340017],accel_mss,speed_ms,0,blend_radius_m)
  speed_ms = 0.005
  movel([-0.230779, -0.945941, -2.745558, -1.020890, 1.570796, 1.340017],accel_mss,speed_ms,0,blend_radius_m)
  speed_ms = 0.025
  movel([-0.232560, -0.948324, -2.744926, -1.019139, 1.570796, 1.338237],accel_mss,speed_ms,0,blend_radius_m)
  movel([-0.232654, -0.948696, -2.744827, -1.018866, 1.570796, 1.338142],accel_mss,speed_ms,0,blend_radius_m)
  movel([-0.232408, -0.949069, -2.744728, -1.018592, 1.570796, 1.338388],accel_mss,speed_ms,0,blend_radius_m)
  movel([-0.230978, -0.949839, -2.744522, -1.018027, 1.570796, 1.339819],accel_mss,speed_ms,0,blend_radius_m)
  movel([-0.224994, -0.951461, -2.744089, -1.016840, 1.570796, 1.345802],accel_mss,speed_ms,0,blend_radius_m)
  movel([-0.216015, -0.953192, -2.743623, -1.015574, 1.570796, 1.354781],accel_mss,speed_ms,0,blend_radius_m)
  movel([-0.205424, -0.955011, -2.743132, -1.014246, 1.570796, 1.365372],accel_mss,speed_ms,0,blend_radius_m)
  movel([-0.184746, -0.958525, -2.742177, -1.011687, 1.570796, 1.386050],accel_mss,speed_ms,0,blend_radius_m)
  movel([-0.173117, -0.960453, -2.741649, -1.010287, 1.570796, 1.397679],accel_mss,speed_ms,0,blend_radius_m)
  movel([-0.172010, -0.960486, -2.741640, -1.010263, 1.570796, 1.398787],accel_mss,speed_ms,0,blend_radius_m)
  movel([-0.170791, -0.960281, -2.741696, -1.010411, 1.570796, 1.400005],accel_mss,speed_ms,0,blend_radius_m)
  movel([-0.169560, -0.959716, -2.741851, -1.010822, 1.570796, 1.401236],accel_mss,speed_ms,0,blend_radius_m)
  movel([-0.168966, -0.959260, -2.741976, -1.011153, 1.570796, 1.401831],accel_mss,speed_ms,0,blend_radius_m)
  movel([-0.168405, -0.958665, -2.742139, -1.011585, 1.570796, 1.402391],accel_mss,speed_ms,0,blend_radius_m)
  movel([-0.167644, -0.957431, -2.742475, -1.012483, 1.570796, 1.403152],accel_mss,speed_ms,0,blend_radius_m)
  movel([-0.167150, -0.956171, -2.742818, -1.013400, 1.570796, 1.403646],accel_mss,speed_ms,0,blend_radius_m)
  movel([-0.165040, -0.949251, -2.744679, -1.018459, 1.570796, 1.405756],accel_mss,speed_ms,0,blend_radius_m)
  movel([-0.163439, -0.942458, -2.746474, -1.023457, 1.570796, 1.407358],accel_mss,speed_ms,0,blend_radius_m)
  movel([-0.162323, -0.935824, -2.748197, -1.028368, 1.570796, 1.408473],accel_mss,speed_ms,0,blend_radius_m)
  movel([-0.161652, -0.929368, -2.749845, -1.033176, 1.570796, 1.409145],accel_mss,speed_ms,0,blend_radius_m)
  movel([-0.161397, -0.923113, -2.751415, -1.037862, 1.570796, 1.409399],accel_mss,speed_ms,0,blend_radius_m)
  movel([-0.161519, -0.917077, -2.752905, -1.042406, 1.570796, 1.409277],accel_mss,speed_ms,0,blend_radius_m)
  movel([-0.161984, -0.911285, -2.754313, -1.046791, 1.570796, 1.408813],accel_mss,speed_ms,0,blend_radius_m)
  movel([-0.162751, -0.905761, -2.755636, -1.050992, 1.570796, 1.408045],accel_mss,speed_ms,0,blend_radius_m)
  movel([-0.163295, -0.903395, -2.756196, -1.052798, 1.570796, 1.407502],accel_mss,speed_ms,0,blend_radius_m)
  movel([-0.164063, -0.901384, -2.756670, -1.054335, 1.570796, 1.406733],accel_mss,speed_ms,0,blend_radius_m)
  movel([-0.165054, -0.899726, -2.757058, -1.055605, 1.570796, 1.405742],accel_mss,speed_ms,0,blend_radius_m)
  movel([-0.166253, -0.898406, -2.757366, -1.056616, 1.570796, 1.404544],accel_mss,speed_ms,0,blend_radius_m)
  movel([-0.167654, -0.897423, -2.757595, -1.057371, 1.570796, 1.403142],accel_mss,speed_ms,0,blend_radius_m)
  movel([-0.169250, -0.896772, -2.757746, -1.057870, 1.570796, 1.401546],accel_mss,speed_ms,0,blend_radius_m)
  movel([-0.171029, -0.896434, -2.757825, -1.058130, 1.570796, 1.399767],accel_mss,speed_ms,0,blend_radius_m)
  movel([-0.172986, -0.896406, -2.757831, -1.058152, 1.570796, 1.397810],accel_mss,speed_ms,0,blend_radius_m)
  movel([-0.175108, -0.896677, -2.757768, -1.057944, 1.570796, 1.395688],accel_mss,speed_ms,0,blend_radius_m)
  movel([-0.177385, -0.897238, -2.757638, -1.057513, 1.570796, 1.393411],accel_mss,speed_ms,0,blend_radius_m)
  movel([-0.179813, -0.898077, -2.757443, -1.056869, 1.570796, 1.390983],accel_mss,speed_ms,0,blend_radius_m)
  movel([-0.182373, -0.899184, -2.757185, -1.056020, 1.570796, 1.388423],accel_mss,speed_ms,0,blend_radius_m)
  movel([-0.187867, -0.902161, -2.756487, -1.053741, 1.570796, 1.382930],accel_mss,speed_ms,0,blend_radius_m)
  movel([-0.193781, -0.906071, -2.755562, -1.050756, 1.570796, 1.377016],accel_mss,speed_ms,0,blend_radius_m)
  movel([-0.199012, -0.910112, -2.754596, -1.047681, 1.570796, 1.371784],accel_mss,speed_ms,0,blend_radius_m)
  movel([-0.204050, -0.914569, -2.753518, -1.044302, 1.570796, 1.366746],accel_mss,speed_ms,0,blend_radius_m)
  movel([-0.208908, -0.919377, -2.752340, -1.040672, 1.570796, 1.361888],accel_mss,speed_ms,0,blend_radius_m)
  movel([-0.213593, -0.924451, -2.751081, -1.036857, 1.570796, 1.357203],accel_mss,speed_ms,0,blend_radius_m)
  movel([-0.218107, -0.929713, -2.749757, -1.032919, 1.570796, 1.352690],accel_mss,speed_ms,0,blend_radius_m)
  movel([-0.222470, -0.935096, -2.748384, -1.028909, 1.570796, 1.348326],accel_mss,speed_ms,0,blend_radius_m)
  movel([-0.230779, -0.945941, -2.745558, -1.020890, 1.570796, 1.340017],accel_mss,speed_ms,0,blend_radius_m)
  movel([-0.232560, -0.948324, -2.744926, -1.019139, 1.570796, 1.338237],accel_mss,speed_ms,0,blend_radius_m)
  movel([-0.232654, -0.948696, -2.744827, -1.018866, 1.570796, 1.338142],accel_mss,speed_ms,0,blend_radius_m)
  movel([-0.232408, -0.949069, -2.744728, -1.018592, 1.570796, 1.338388],accel_mss,speed_ms,0,blend_radius_m)
  movel([-0.231956, -0.949314, -2.744662, -1.018412, 1.570796, 1.338841],accel_mss,speed_ms,0,blend_radius_m)
  speed_ms = 0.005
  movel([-0.231956, -0.940618, -2.738783, -1.032988, 1.570796, 1.338841],accel_mss,speed_ms,0,blend_radius_m)
  speed_ms = 0.040
  movel([-0.253357, -0.923350, -2.743246, -1.045793, 1.570796, 1.317439],accel_mss,speed_ms,0,blend_radius_m)
  speed_ms = 0.005
  movel([-0.253357, -0.931954, -2.749188, -1.031247, 1.570796, 1.317439],accel_mss,speed_ms,0,blend_radius_m)
  speed_ms = 0.025
  movel([-0.253972, -0.929944, -2.749699, -1.032746, 1.570796, 1.316825],accel_mss,speed_ms,0,blend_radius_m)
  movel([-0.254986, -0.928294, -2.750116, -1.033979, 1.570796, 1.315810],accel_mss,speed_ms,0,blend_radius_m)
  movel([-0.256378, -0.927047, -2.750430, -1.034911, 1.570796, 1.314418],accel_mss,speed_ms,0,blend_radius_m)
  movel([-0.258113, -0.926231, -2.750635, -1.035523, 1.570796, 1.312683],accel_mss,speed_ms,0,blend_radius_m)
  movel([-0.263111, -0.925308, -2.750867, -1.036214, 1.570796, 1.307685],accel_mss,speed_ms,0,blend_radius_m)
  movel([-0.264380, -0.924829, -2.750987, -1.036573, 1.570796, 1.306417],accel_mss,speed_ms,0,blend_radius_m)
  movel([-0.265348, -0.924129, -2.751161, -1.037098, 1.570796, 1.305449],accel_mss,speed_ms,0,blend_radius_m)
  movel([-0.265864, -0.923156, -2.751404, -1.037829, 1.570796, 1.304932],accel_mss,speed_ms,0,blend_radius_m)
  movel([-0.265771, -0.921839, -2.751731, -1.038819, 1.570796, 1.305025],accel_mss,speed_ms,0,blend_radius_m)
  movel([-0.264993, -0.920087, -2.752165, -1.040137, 1.570796, 1.305804],accel_mss,speed_ms,0,blend_radius_m)
  movel([-0.263876, -0.918672, -2.752514, -1.041203, 1.570796, 1.306920],accel_mss,speed_ms,0,blend_radius_m)
  movel([-0.262511, -0.917555, -2.752788, -1.042046, 1.570796, 1.308286],accel_mss,speed_ms,0,blend_radius_m)
  movel([-0.260997, -0.916704, -2.752997, -1.042688, 1.570796, 1.309799],accel_mss,speed_ms,0,blend_radius_m)
  movel([-0.257929, -0.915673, -2.753249, -1.043467, 1.570796, 1.312867],accel_mss,speed_ms,0,blend_radius_m)
  movel([-0.255441, -0.915296, -2.753341, -1.043752, 1.570796, 1.315355],accel_mss,speed_ms,0,blend_radius_m)
  movel([-0.256857, -0.913320, -2.753821, -1.045248, 1.570796, 1.313940],accel_mss,speed_ms,0,blend_radius_m)
  movel([-0.258716, -0.911912, -2.754162, -1.046315, 1.570796, 1.312080],accel_mss,speed_ms,0,blend_radius_m)
  movel([-0.263245, -0.910104, -2.754598, -1.047688, 1.570796, 1.307552],accel_mss,speed_ms,0,blend_radius_m)
  movel([-0.267977, -0.908443, -2.754996, -1.048950, 1.570796, 1.302820],accel_mss,speed_ms,0,blend_radius_m)
  movel([-0.270097, -0.907216, -2.755289, -1.049883, 1.570796, 1.300699],accel_mss,speed_ms,0,blend_radius_m)
  movel([-0.271870, -0.905477, -2.755703, -1.051209, 1.570796, 1.298926],accel_mss,speed_ms,0,blend_radius_m)
  movel([-0.272742, -0.904111, -2.756027, -1.052251, 1.570796, 1.298054],accel_mss,speed_ms,0,blend_radius_m)
  movel([-0.273247, -0.902815, -2.756333, -1.053241, 1.570796, 1.297549],accel_mss,speed_ms,0,blend_radius_m)
  movel([-0.273420, -0.901595, -2.756620, -1.054174, 1.570796, 1.297376],accel_mss,speed_ms,0,blend_radius_m)
  movel([-0.273287, -0.900461, -2.756886, -1.055042, 1.570796, 1.297509],accel_mss,speed_ms,0,blend_radius_m)
  movel([-0.272891, -0.899428, -2.757128, -1.055833, 1.570796, 1.297905],accel_mss,speed_ms,0,blend_radius_m)
  movel([-0.272260, -0.898496, -2.757346, -1.056548, 1.570796, 1.298536],accel_mss,speed_ms,0,blend_radius_m)
  movel([-0.271436, -0.897683, -2.757535, -1.057171, 1.570796, 1.299360],accel_mss,speed_ms,0,blend_radius_m)
  movel([-0.270446, -0.896996, -2.757694, -1.057699, 1.570796, 1.300351],accel_mss,speed_ms,0,blend_radius_m)
  movel([-0.269329, -0.896446, -2.757822, -1.058121, 1.570796, 1.301467],accel_mss,speed_ms,0,blend_radius_m)
  movel([-0.268126, -0.896047, -2.757914, -1.058427, 1.570796, 1.302670],accel_mss,speed_ms,0,blend_radius_m)
  movel([-0.265587, -0.895732, -2.757987, -1.058669, 1.570796, 1.305209],accel_mss,speed_ms,0,blend_radius_m)
  movel([-0.263116, -0.896130, -2.757895, -1.058364, 1.570796, 1.307680],accel_mss,speed_ms,0,blend_radius_m)
  movel([-0.260996, -0.897318, -2.757619, -1.057451, 1.570796, 1.309800],accel_mss,speed_ms,0,blend_radius_m)
  movel([-0.261112, -0.894740, -2.758216, -1.059433, 1.570796, 1.309684],accel_mss,speed_ms,0,blend_radius_m)
  movel([-0.261559, -0.892556, -2.758719, -1.061115, 1.570796, 1.309237],accel_mss,speed_ms,0,blend_radius_m)
  movel([-0.262267, -0.890682, -2.759147, -1.062560, 1.570796, 1.308529],accel_mss,speed_ms,0,blend_radius_m)
  movel([-0.265217, -0.885894, -2.760232, -1.066263, 1.570796, 1.305579],accel_mss,speed_ms,0,blend_radius_m)
  movel([-0.267134, -0.882394, -2.761017, -1.068978, 1.570796, 1.303662],accel_mss,speed_ms,0,blend_radius_m)
  movel([-0.267684, -0.880727, -2.761388, -1.070275, 1.570796, 1.303113],accel_mss,speed_ms,0,blend_radius_m)
  movel([-0.267937, -0.879096, -2.761749, -1.071544, 1.570796, 1.302860],accel_mss,speed_ms,0,blend_radius_m)
  movel([-0.267925, -0.877533, -2.762094, -1.072762, 1.570796, 1.302871],accel_mss,speed_ms,0,blend_radius_m)
  movel([-0.267674, -0.876057, -2.762418, -1.073914, 1.570796, 1.303122],accel_mss,speed_ms,0,blend_radius_m)
  movel([-0.267218, -0.874693, -2.762716, -1.074980, 1.570796, 1.303578],accel_mss,speed_ms,0,blend_radius_m)
  movel([-0.266583, -0.873460, -2.762985, -1.075944, 1.570796, 1.304213],accel_mss,speed_ms,0,blend_radius_m)
  movel([-0.265800, -0.872385, -2.763218, -1.076786, 1.570796, 1.304996],accel_mss,speed_ms,0,blend_radius_m)
  movel([-0.264899, -0.871492, -2.763412, -1.077485, 1.570796, 1.305897],accel_mss,speed_ms,0,blend_radius_m)
  movel([-0.263912, -0.870806, -2.763560, -1.078023, 1.570796, 1.306885],accel_mss,speed_ms,0,blend_radius_m)
  movel([-0.262870, -0.870349, -2.763659, -1.078381, 1.570796, 1.307926],accel_mss,speed_ms,0,blend_radius_m)
  movel([-0.261802, -0.870144, -2.763703, -1.078542, 1.570796, 1.308994],accel_mss,speed_ms,0,blend_radius_m)
  movel([-0.260739, -0.870218, -2.763687, -1.078484, 1.570796, 1.310058],accel_mss,speed_ms,0,blend_radius_m)
  movel([-0.259716, -0.870596, -2.763606, -1.078187, 1.570796, 1.311080],accel_mss,speed_ms,0,blend_radius_m)
  movel([-0.258762, -0.871299, -2.763454, -1.077636, 1.570796, 1.312035],accel_mss,speed_ms,0,blend_radius_m)
  movel([-0.257907, -0.872351, -2.763226, -1.076812, 1.570796, 1.312889],accel_mss,speed_ms,0,blend_radius_m)
  movel([-0.257181, -0.873767, -2.762918, -1.075704, 1.570796, 1.313616],accel_mss,speed_ms,0,blend_radius_m)
  movel([-0.256154, -0.870916, -2.763536, -1.077936, 1.570796, 1.314643],accel_mss,speed_ms,0,blend_radius_m)
  movel([-0.255439, -0.868208, -2.764119, -1.080062, 1.570796, 1.315357],accel_mss,speed_ms,0,blend_radius_m)
  movel([-0.254976, -0.865614, -2.764673, -1.082101, 1.570796, 1.315820],accel_mss,speed_ms,0,blend_radius_m)
  movel([-0.254699, -0.863105, -2.765206, -1.084079, 1.570796, 1.316097],accel_mss,speed_ms,0,blend_radius_m)
  movel([-0.254108, -0.853296, -2.767251, -1.091842, 1.570796, 1.316688],accel_mss,speed_ms,0,blend_radius_m)
  movel([-0.253785, -0.849611, -2.768005, -1.094773, 1.570796, 1.317011],accel_mss,speed_ms,0,blend_radius_m)
  movel([-0.252996, -0.845027, -2.768931, -1.098431, 1.570796, 1.317800],accel_mss,speed_ms,0,blend_radius_m)
  movel([-0.252214, -0.842644, -2.769408, -1.100337, 1.570796, 1.318583],accel_mss,speed_ms,0,blend_radius_m)
